(* IEC 61131-3 sources: daoli-st-library/DL_Process (part 46) *)

(* ---- FB_DL_PowderDosingLoss.st ---- *)
// =====================================================================
// FB_DL_PowderDosingLoss.st
// 粉料失重秤增量式配料（皮重→粗给/慢给→落差补偿→稳定结算→学习）
// Loss-in-weight powder dosing FB
// 码位: 16#0005_0458 ~ 16#0005_045C (本件独占 5 槽)
// 修改记录: R29 初版 (按 DISPATCH_R29 序 18)
// =====================================================================
FUNCTION_BLOCK FB_DL_PowderDosingLoss
VAR_INPUT
    bEnable      : BOOL  := FALSE;    // 使能 / Enable
    bStart       : BOOL  := FALSE;    // 上升沿开始一批 / Start batch on edge
    bReset       : BOOL  := FALSE;    // 复位 / Reset
    fWeight_g    : REAL  := 0.0;      // 秤读数 0~500000 g / Scale weight [g]
    fTarget_g    : REAL  := 1000.0;   // 目标投料量 >0 g / Target dose [g]
    fTare_g      : REAL  := 0.0;      // 皮重 ≥0 g / Tare [g]
    fSlowBand_g  : REAL  := 100.0;    // 转慢速余量 >0 g / Slow-down band [g]
    fLead_g      : REAL  := 0.0;      // 落差学习初值 0~500 g / Lead compensation [g]
    fLeadMax_g   : REAL  := 300.0;    // 落差限幅 1~2000 g / Lead limit [g]
    fDevMax_g    : REAL  := 5.0;      // 允许偏差 >0 g / Allowed deviation [g]
    bSlowCmd     : BOOL  := FALSE;    // 慢速输出确认 / Slow feed ack
    tSettleTime  : TIME  := T#500MS;  // 停料稳定时 T#10MS~T#10S / Settle time [s]
    tBatchMax    : TIME  := T#2M;     // 单批超时 T#1S~T#30M / Batch timeout [s]
END_VAR
VAR_OUTPUT
    fNet_g       : REAL;              // 本批净投料 g / Net dosed [g]
    fErr_g       : REAL;              // 本批偏差 g / Deviation [g]
    bDone        : BOOL;              // 批完成（单拍）/ Batch done pulse
    bBusy        : BOOL;              // 配料中 / Busy
    fLeadLearn_g : REAL;              // 更新后落差学习值 g / Learned lead [g]
    eErr         : UDINT;             // 错误码 / Error code
END_VAR
VAR
    rtrigStart   : R_TRIG;            // 启动沿检测（无条件刷新）/ Start edge detector
    tonSettle    : TON;               // 停料稳定定时器（无条件刷新）/ Settle timer
    tonBatch     : TON;               // 单批超时定时器（无条件刷新）/ Batch timeout timer
    fTareSnap_g  : REAL;              // 批开始皮重快照 / Tare snapshot at batch start [g]
    fWeightPrev  : REAL;              // 上拍秤读数快照 / Previous weight snapshot [g]
    fNetNow_g    : REAL;              // 本拍净重 / Net weight this cycle [g]
    fNetStart_g  : REAL;              // 批开始净重基准 / Net baseline at batch start [g]
    fStopPt_g    : REAL;              // 提前停止点（目标-慢带-落差）/ Early stop point [g]
    bFastPhase   : BOOL;              // 高速给料相 / Fast feed phase
    bSettling    : BOOL;              // 停料稳定相 / Settling phase
    tSettleS     : REAL;              // 稳定时秒值 / Settle seconds [s]
    tBatchMaxS   : REAL;              // 批超时秒值 / Batch timeout seconds [s]
    bAbortLatch  : BOOL := FALSE;     // 中止锁存（方向反/超时）/ Abort latch
    xFirstScan   : BOOL  := TRUE;     // 首扫标记 / First-scan flag
END_VAR

// ---------------------------------------------------------------------
// 代码位表（本件独占，勿复用）:
//   16#0005_0458 信息 批完成、偏差在容差内
//   16#0005_0459 故障 秤值非有限 / 皮重为负或超量程 / tSettleTime 非法
//   16#0005_045A 故障 fTarget_g ≤ 0 / fSlowBand_g ≥ fTarget_g / fLeadMax_g ≤ 0（组态错）
//   16#0005_045B 信息 批完成但偏差 > fDevMax_g → 结算照出、落差不学习
//   16#0005_045C 故障 进料期重量上升（方向反）或超 tBatchMax → 中止锁存（方向反优先）
// ---------------------------------------------------------------------

// ---- 时间转秒 / Times to seconds ----
tSettleS := TIME_TO_REAL(tSettleTime) / 1000.0;     // 稳定时秒 / Settle [s]
tBatchMaxS := TIME_TO_REAL(tBatchMax) / 1000.0;     // 批超时秒 / Batch max [s]

// ---- 启动沿检测（无条件刷新）/ Start edge, unconditional ----
rtrigStart(CLK := bStart);      // 沿检测 / Edge detection

// ---- 非有限与皮重闸（故障级）/ Finite and tare gate ----
IF (fWeight_g <> fWeight_g) OR (ABS(fWeight_g) >= 1.0E12)
   OR (fTare_g < 0.0) OR (fTare_g > 500000.0)
   OR (tSettleTime = T#0MS) OR (tSettleS < 0.01) OR (tSettleS > 10.0) THEN
    bBusy := FALSE;             // 停止 / Not busy
    bAbortLatch := TRUE;        // 中止锁存 / Abort latch
    eErr := 16#0005_0459;       // 故障码 / Fault code
    RETURN;                     // 本拍结束 / End of cycle
END_IF

// ---- 组态错闸 / Configuration fault gate ----
IF (fTarget_g <= 0.0) OR (fSlowBand_g >= fTarget_g) OR (fLeadMax_g <= 0.0)
   OR (fDevMax_g <= 0.0)
   OR (tBatchMax = T#0MS) OR (tBatchMaxS < 1.0) OR (tBatchMaxS > 1800.0) THEN
    eErr := 16#0005_045A;       // 故障码 / Fault code
    RETURN;                     // 本拍结束 / End of cycle
END_IF

// ---- 首扫初始化（R16 首扫纪律）/ First-scan initialization ----
IF xFirstScan THEN
    fLeadLearn_g := fLead_g;    // 学习值取初值 / Learn value from init
    fWeightPrev := fWeight_g;   // 快照对齐 / Snapshot align
    bDone := FALSE;             // 脉冲复位 / Pulse reset
    xFirstScan := FALSE;        // 清标记 / Clear flag
END_IF

// ---- 完成脉冲单拍化 / Done pulse one-cycle ----
IF bDone THEN
    bDone := FALSE;             // 下一拍清 / Clear next cycle
END_IF

// ---- 使能撤销 / Disable ----
IF NOT bEnable THEN
    bBusy := FALSE;             // 停止 / Not busy
    bFastPhase := FALSE;        // 粗给退出 / Fast off
    bSettling := FALSE;         // 稳定退出 / Settle off
    eErr := 16#0005_0458;       // 信息级：空闲 / Info: idle
    RETURN;                     // 本拍结束 / End of cycle
END_IF

// ---- 复位：清中止锁存与学习值回初值 / Reset: clear latch, learn back to init ----
IF bReset THEN
    bAbortLatch := FALSE;       // 解锁存 / Release latch
    bBusy := FALSE;             // 停止 / Not busy
    bFastPhase := FALSE;        // 粗给退出 / Fast off
    bSettling := FALSE;         // 稳定退出 / Settle off
    fLeadLearn_g := fLead_g;    // 学习值回初值 / Learn to init
END_IF

// ---- 中止锁存路径 / Abort latch path ----
IF bAbortLatch THEN
    bBusy := FALSE;             // 停止（保留已投量）/ Stopped, dose kept
    eErr := 16#0005_045C;       // 故障码回放 / Fault code replay
    RETURN;                     // 本拍结束 / End of cycle
END_IF

// ---- 每拍净重与方向监控 / Per-cycle net and direction monitor ----
fNetNow_g := fWeight_g - fTare_g;   // 净重 / Net [g]
IF fNetNow_g < 0.0 THEN
    fNetNow_g := 0.0;           // 负值钳 0 / Clamp to 0
    eErr := 16#0005_0459;       // 槽 2 登记 / Slot 2
END_IF

// ---- 启动沿受理（bBusy=FALSE 才受理）/ Accept start edge when idle ----
IF rtrigStart.Q AND (NOT bBusy) THEN
    fTareSnap_g := fTare_g;     // 皮重快照 / Tare snapshot
    fNetStart_g := fNetNow_g;   // 净重基准 / Net baseline
    fWeightPrev := fWeight_g;   // 快照对齐 / Snapshot align
    fStopPt_g := fTarget_g - fSlowBand_g - fLeadLearn_g;    // 提前停止点含落差 / Stop point with lead
    IF fStopPt_g < 0.0 THEN
        fStopPt_g := 0.0;       // 防负停止点 / Guard negative stop
    END_IF
    bBusy := TRUE;              // 配料中 / Busy
    bFastPhase := TRUE;         // 粗给开始 / Fast feed
    bSettling := FALSE;         // 非稳定相 / Not settling
END_IF

// ---- 批运行路径 / Batch active path ----
IF bBusy THEN
    // 单批超时监控 / Batch timeout monitor
    tonBatch(IN := bBusy, PT := tBatchMax);     // 无条件刷新 / Unconditional refresh

    // 方向监控：进料期重量上升 → 方向反（根因优先，先于超时判）/ Direction: rising weight fault first
    IF fWeight_g > (fWeightPrev + 1.0) THEN
        bAbortLatch := TRUE;    // 中止锁存 / Abort latch
        bBusy := FALSE;         // 停止 / Not busy
        bFastPhase := FALSE;    // 粗给退出 / Fast off
        bSettling := FALSE;     // 稳定退出 / Settle off
        eErr := 16#0005_045C;   // 故障码：方向反 / Fault code: reversed
        fWeightPrev := fWeight_g;   // 快照对齐 / Align snapshot
        RETURN;                 // 本拍结束 / End of cycle
    END_IF

    // 批超时（方向反已优先返回）/ Batch timeout after direction check
    IF tonBatch.Q THEN
        bAbortLatch := TRUE;    // 中止锁存 / Abort latch
        bBusy := FALSE;         // 停止（保留已投量）/ Stopped, dose kept
        bFastPhase := FALSE;    // 粗给退出 / Fast off
        bSettling := FALSE;     // 稳定退出 / Settle off
        eErr := 16#0005_045C;   // 故障码：超时 / Fault code: timeout
        RETURN;                 // 本拍结束 / End of cycle
    END_IF

    // ---- 给料相控制 / Feed phase control ----
    IF bFastPhase THEN
        // 高速粗给：净投量未达提前停止点 / Fast: below stop point
        IF (fNetNow_g - fNetStart_g) >= fStopPt_g THEN
            bFastPhase := FALSE;    // 转慢速精给 / To slow feed
        END_IF
        // 慢速转换确认（bSlowCmd 为外部确认，此处登记不强制）/ Slow ack registered externally
    END_IF

    // 停料判定：慢给相已达目标（含落差提前）/ Stop: reached target with lead
    IF (NOT bFastPhase) AND ((fNetNow_g - fNetStart_g) >= (fTarget_g - fLeadLearn_g)) THEN
        bSettling := TRUE;      // 停料稳定相 / Settling
        tonSettle(IN := TRUE, PT := tSettleTime);   // 稳定计时 / Settle timing
    END_IF

    // ---- 稳定后结算 / Settle then finalize ----
    IF bSettling THEN
        tonSettle(IN := TRUE, PT := tSettleTime);   // 无条件刷新 / Unconditional refresh
        IF tonSettle.Q THEN
            fNet_g := fNetNow_g - fNetStart_g;  // 结算净投量 / Finalize net
            fErr_g := fNet_g - fTarget_g;       // 偏差 / Deviation
            bDone := TRUE;      // 完成脉冲 / Done pulse
            bBusy := FALSE;     // 停止 / Not busy
            bSettling := FALSE; // 稳定退出 / Settle off
            IF ABS(fErr_g) <= fDevMax_g THEN
                // 落差学习：LIMIT(0, fLead + 0.5×fErr, fLeadMax)，0.5 阻尼防振荡
                // Lead learning: LIMIT with 0.5 damping factor
                fLeadLearn_g := fLeadLearn_g + 0.5 * fErr_g;    // 学习更新 / Learn update
                IF fLeadLearn_g < 0.0 THEN
                    fLeadLearn_g := 0.0;    // 下限 / Lower limit
                ELSIF fLeadLearn_g > fLeadMax_g THEN
                    fLeadLearn_g := fLeadMax_g;     // 上限 / Upper limit
                END_IF
                eErr := 16#0005_0458;   // 信息级：批完成 / Info: done
            ELSE
                eErr := 16#0005_045B;   // 信息级：超差结算不学习 / Info: no learning
            END_IF
        END_IF
    END_IF
ELSE
    tonBatch(IN := FALSE, PT := tBatchMax);     // 定时器复位 / Timer reset
    tonSettle(IN := FALSE, PT := tSettleTime);  // 定时器复位 / Timer reset
END_IF

// ---- 上拍快照更新 / Previous snapshot update ----
fWeightPrev := fWeight_g;       // 快照 / Snapshot

END_FUNCTION_BLOCK

(* ---- FB_DL_PressFitCurveArchive.st ---- *)
(*
  Component : FB_DL_PressFitCurveArchive
  Category  : DL_Process
  Type      : FB
  Version   : 1.0.0
  CodeSeg   : 16#06_0_3B
  Summary   : 压装曲线特征点归档与批次追溯：四特征点环形缓存按批次号索引，R_TRIG 沿触发归档。
              Press-fit curve feature archive by batch index in a ring buffer, triggered on a rising edge.
  溯源声明  : 道莅自研 clean-room
  边界安全  : 批次号域闸（> 0，防非法索引）；环形缓冲下标 1..NMAX 硬界，写前钳制防越界；
              特征点非有限（NaN 自反 + Inf 上限）拦截；查询命中用整数相等（DINT）；
              R_TRIG 每拍无条件刷新（段 0）；缓冲满环回写并置 bWrapped 提示；计数防回卷。
  复用      : 无
*)

FUNCTION_BLOCK FB_DL_PressFitCurveArchive
VAR_INPUT
    bRun       : BOOL;                  (* 归档使能 · Enable *)
    bArchCmd   : BOOL;                  (* 归档指令 [事件]，沿触发 · Archive command, edge *)
    nBatchNo   : DINT;                  (* 批次号 [号]，域 > 0 · Batch number *)
    fF1KN      : LREAL;                 (* 特征点 1：起步压力 [kN] · Feature 1 onset force *)
    fF2MM      : LREAL;                 (* 特征点 2：起步位移 [mm] · Feature 2 onset travel *)
    fF3KN      : LREAL;                 (* 特征点 3：峰值压力 [kN] · Feature 3 peak force *)
    fF4MM      : LREAL;                 (* 特征点 4：终点位移 [mm] · Feature 4 end travel *)
    nQueryNo   : DINT;                  (* 追溯查询批次号 [号] · Query batch number *)
    fEps       : LREAL := 1.0E-6;       (* 浮点判零容差 [实数域] · Floating zero tolerance *)
END_VAR
VAR_OUTPUT
    bArchOk  : BOOL;                    (* 本拍归档成功 [开关] · Archive succeeded this scan *)
    bWrapped : BOOL;                    (* 环已回卷覆盖标志 · Ring wrapped flag *)
    bFound   : BOOL;                    (* 查询命中标志 · Query hit flag *)
    fQ1KN    : LREAL;                   (* 查询特征 1 [kN] · Queried feature 1 *)
    fQ2MM    : LREAL;                   (* 查询特征 2 [mm] · Queried feature 2 *)
    fQ3KN    : LREAL;                   (* 查询特征 3 [kN] · Queried feature 3 *)
    fQ4MM    : LREAL;                   (* 查询特征 4 [mm] · Queried feature 4 *)
    nUsed    : INT;                     (* 环内已用槽数 [槽] · Used slots *)
    bError   : BOOL;                    (* 故障标志，与故障码配对 · Fault flag paired with codes *)
    uErrorId : UDINT;                   (* 事件码 16#0000_003B，0 无事件 · Event code *)
END_VAR
VAR
    uCode   : WORD;     (* 码位暂存，每拍重算 [码] · Code staging *)
    rTrigArc: R_TRIG;   (* 归档上升沿，每拍无条件刷新 · Archive edge detection *)
    aIdx    : ARRAY[1..8] OF DINT;      (* 批次号索引槽 [号] · Batch index slots *)
    aF1     : ARRAY[1..8] OF LREAL;     (* 特征 1 缓存 [kN] · Feature 1 buffer *)
    aF2     : ARRAY[1..8] OF LREAL;     (* 特征 2 缓存 [mm] · Feature 2 buffer *)
    aF3     : ARRAY[1..8] OF LREAL;     (* 特征 3 缓存 [kN] · Feature 3 buffer *)
    aF4     : ARRAY[1..8] OF LREAL;     (* 特征 4 缓存 [mm] · Feature 4 buffer *)
    nHead   : INT;      (* 环形写头下标 [索引] · Ring head index *)
    nI      : INT;      (* 查询循环下标 [索引] · Query loop index *)
    bSigOk  : BOOL;     (* 输入有效标志 · Input validity flag *)
    nCycles : UDINT;    (* 归档累计 [次]，防回卷 · Archive count *)
END_VAR
VAR CONSTANT
    DL_PCA_NMAX : INT := 8;             (* 环形缓冲容量 [槽] · Ring capacity *)
    DL_PCA_WRAP : UDINT := 4294967290;  (* 计数防回卷余量 [次] · Counter wrap guard *)
END_VAR

(* === 段 0 · 实例刷新（每拍无条件，红线 7）=== *)
IF nHead < 1 THEN
    nHead := 1;                         (* 写头初值钳 1，防数组零下标越界 / Clamp the head to one *)
END_IF
rTrigArc(CLK := bArchCmd);              (* 归档沿检测 / Archive edge *)

(* === 段 1 · 输入校验与量程闸 === *)
uCode := 16#0000;                       // 每拍清码（可达清零基线）/ Clear codes each scan
bSigOk := (nBatchNo > 0)                                             // 批次号正域闸 / Batch number gate
          AND (fF1KN = fF1KN) AND (fF2MM = fF2MM)                     // 特征点非有限拦截 / Non-finite guards
          AND (fF3KN = fF3KN) AND (fF4MM = fF4MM)
          AND (ABS(fF1KN) < 1.0E308) AND (ABS(fF3KN) < 1.0E308)       // Inf 上限判据 / Inf limits
          AND (ABS(fF2MM) < 1.0E308) AND (ABS(fF4MM) < 1.0E308)
          AND (fF3KN > fF1KN);                                        // 峰值起步序闸 / Peak above onset
IF NOT bSigOk THEN
    uCode := 16#003B;                   // 故障级：域外，归档拒绝 / Fault: domain invalid
END_IF

(* === 段 2 · 主逻辑：环形归档与批次追溯 === *)
bArchOk := FALSE;                       (* 归档成功标志单拍重建 / Rebuild the success flag *)
IF rTrigArc.Q AND bRun THEN
    IF bSigOk THEN
        aIdx[nHead] := nBatchNo;        (* 写批次索引（头下标受 NMAX 硬界）/ Write the index *)
        aF1[nHead] := fF1KN;            (* 写特征 1 [kN] / Write feature 1 *)
        aF2[nHead] := fF2MM;            (* 写特征 2 [mm] / Write feature 2 *)
        aF3[nHead] := fF3KN;            (* 写特征 3 [kN] / Write feature 3 *)
        aF4[nHead] := fF4MM;            (* 写特征 4 [mm] / Write feature 4 *)
        bArchOk := TRUE;                (* 归档成功 / Archive done *)
        IF nUsed < DL_PCA_NMAX THEN
            nUsed := nUsed + 1;         (* 未满先增用量 / Grow usage *)
        ELSE
            bWrapped := TRUE;           (* 满环回卷提示 / Ring wrapped flag *)
        END_IF
        nHead := (nHead MOD DL_PCA_NMAX) + 1;   (* 写头循环推进，界内 / Advance the head in bounds *)
        IF nCycles < DL_PCA_WRAP THEN
            nCycles := nCycles + 1;     (* 归档计数 / Count archives *)
        END_IF
    END_IF
END_IF
(* 追溯查询：按批次号线性匹配（DINT 等值合法）/ Trace query by batch number *)
bFound := FALSE;                        (* 命中标志单拍重建 / Rebuild the hit flag *)
IF (nQueryNo > 0) AND (nUsed >= 1) THEN
    FOR nI := 1 TO DL_PCA_NMAX DO
        IF nI <= nUsed THEN
            IF aIdx[nI] = nQueryNo THEN
                fQ1KN := aF1[nI];       (* 命中回放特征 1 [kN] / Replay feature 1 *)
                fQ2MM := aF2[nI];       (* 回放特征 2 [mm] / Replay feature 2 *)
                fQ3KN := aF3[nI];       (* 回放特征 3 [kN] / Replay feature 3 *)
                fQ4MM := aF4[nI];       (* 回放特征 4 [mm] / Replay feature 4 *)
                bFound := TRUE;         (* 命中 / Hit *)
                EXIT;                   (* 单命中即止 / Stop on first hit *)
            END_IF
        END_IF
    END_FOR
END_IF

(* === 段 3 · 输出映射与故障码 === *)
IF NOT bFound THEN
    fQ1KN := 0.0;                       (* 未命中输出安全零（哨兵）/ Safe zeros on miss *)
    fQ2MM := 0.0;
    fQ3KN := 0.0;
    fQ4MM := 0.0;
END_IF
IF NOT bRun THEN
    bWrapped := FALSE;                  (* 撤使能清回卷提示（可达清零）/ Clear on disable *)
END_IF
bError := (uCode <> 16#0000);           (* 故障标志配对 / Fault flag paired *)
uErrorId := WORD_TO_UDINT(uCode);       (* 码位单点写入（16#0000_003B 形态）/ Single write point *)
END_FUNCTION_BLOCK

(* ---- FB_DL_PrintRegisterAutoTrimSeq.st ---- *)
(*
  DL Factory R83 | FB_DL_PrintRegisterAutoTrimSeq
  功能：印刷套准自动调整状态机，横纵套准误差超差后按三级阶梯逐级小步修正，每步等稳定窗后复评，超步数上限锁故障码。
  开源溯源：无（clean-room 自研，依据公开工艺公式，来源=行业通用公式，许可证=MIT，借鉴点=公式结构）
  规则：R1-R21 全遵守
  ------------------------------------------------------------------
  分类 DL_Process ｜ 复杂度 cx4 ｜ 版本 v1.0.0 ｜ 平台 纯 IEC 61131-3（TON、R_TRIG、LREAL）
  边界：一 只出三级修正命令，不驱动版辊电机本体、不做套准标记识别（识别归前级视觉件属主）；
        二 阶梯次序固定：一 色标偏移（管横向）→ 二 版辊相位（管纵向）→ 三 张力微调（管纵向残差）；
           一与二同属偏移域共用 eVern 相、由 _nLadder 区分下发通道；三独立占 eTens 相（力值量禁与长度量混加）；
        三 每步下发后等回执沿（脉冲语义，须回零后再置位），否则超时锁 104；每相只允许一个专属定时器，
           IN 只串本相使能与锁存闸，相迁移即 IN 归假并自复位（R18）；tonVern 与 tonTens 分属互斥相、
           无同拍双窗，故 R100 配比约束不适用；
        四 小步下发前方向分列（偏正 ｜ 偏负各占一分支，R146），下发后立即饱和到本通道限值；
        五 命令累加量在复位沿保持末值（已下发修正不得被复位抹掉），作用域在段 1 逐项声明；
           无全局变量、无外部变量声明、无物理地址寻址。
  量纲自检：长度量 [mm] 通道 = fErrCross / fTolCross / fStepVernier / fCmdLimit 与 fErrMachine / fTolMachine / fStepPhase；
        力值量 [N] 通道 = fStepTension / fTensLimit（禁与长度量相加）；组态闸另校各步长落在本通道限值内防越窗振荡。
  输出契约：三级命令为累加型且已饱和；bDone 为电平保持位（新循环起点同拍清零，R28 5.9）；iErrCode 为锁存回放，故障锁存唯一解除路径为 bReset 上升沿（R188）。
  修订记录：2026-11-24 v1.0.0 R83 首版（批 R83 · 序号 37）
*)

TYPE E_DL_PraPhase :
(
    eIdle   := 0,  // 空闲等启动沿 / idle, waiting for the start edge
    eEval   := 10, // 评估：判容差选阶梯并下发（单拍相）/ evaluate, judge and issue in one scan
    eVern   := 20, // 偏移修正等回执（承载阶梯一二）/ offset trim, waiting for the acknowledgement
    eTens   := 30, // 张力修正等回执（承载阶梯三）/ tension trim, waiting for the acknowledgement
    eSettle := 40, // 稳定等稳定窗 / settling, waiting for the window
    eDone   := 50, // 完成：误差在容差内 / done, the error is inside the tolerance
    eFault  := 90  // 故障：成因锁存等复位沿 / fault, the cause is latched until the reset edge
);
END_TYPE

TYPE E_DL_PraCause :
(
    eNone      := 0, // 无成因 / no cause
    eCfgBad    := 1, // 组态越域或量纲失配（故障级，与 bError 配对）/ configuration out of domain, fault grade paired with bError
    eNotFinite := 2, // 入参非有限 NaN 或 Inf（故障级，与 bError 配对）/ non-finite input, fault grade paired with bError
    eStepLimit := 3, // 步数上限耗尽仍超差（故障级，与 bError 配对）/ step budget exhausted, fault grade paired with bError
    eAckTo     := 4, // 步进回执超时（故障级，与 bError 配对）/ acknowledgement timeout, fault grade paired with bError
    ePhaseBad  := 5  // 非法相位兜底（故障级，与 bError 配对）/ illegal phase fallback, fault grade paired with bError
);
END_TYPE

FUNCTION_BLOCK FB_DL_PrintRegisterAutoTrimSeq
VAR CONSTANT
    DL_PRA_LADDER_VERN   : INT := 1; // 阶梯一：色标偏移通道 [级] / ladder one, the register mark offset channel [stage]
    DL_PRA_LADDER_PHASE  : INT := 2; // 阶梯二：版辊相位通道 [级] / ladder two, the plate cylinder phase channel [stage]
    DL_PRA_LADDER_TENS   : INT := 3; // 阶梯三：张力微调通道 [级] / ladder three, the tension trim channel [stage]
    DL_PRA_PHASE_TRY_MAX : INT := 2; // 阶梯二连续复用预算，超限升阶梯三 [次] / the reuse budget of ladder two [time]
END_VAR
VAR_INPUT
    bEnable      : BOOL := TRUE;   // 使能，失能退回空闲（命令保持末值）[-] / enable, a disable returns to idle holding the commands
    bReset       : BOOL := FALSE;  // 复位上升沿清故障锁存与步数 [-]/ reset rising edge clears the latch and the steps
    bStart       : BOOL := FALSE;  // 启动电平，上升沿起一轮调整 [-]/ start level, its rising edge begins one round
    bStepAck     : BOOL := FALSE;  // 步进执行回执（脉冲语义须回零）[-]/ the step acknowledgement, pulse semantics
    fErrCross    : LREAL := 0.0;   // 横向套准误差（正 = 偏大）[mm] / the cross register error, positive means too large [mm]
    fErrMachine  : LREAL := 0.0;   // 纵向套准误差（正 = 偏大）[mm] / the machine register error, positive means too large [mm]
    fTolCross    : LREAL := 0.10;  // 横向容差半带宽 [mm] / the cross tolerance half band [mm]
    fTolMachine  : LREAL := 0.10;  // 纵向容差半带宽 [mm] / the machine tolerance half band [mm]
    fStepVernier : LREAL := 0.05;  // 色标偏移单步量（阶梯一）[mm] / the offset step of ladder one [mm]
    fStepPhase   : LREAL := 0.05;  // 版辊相位单步等效位移（阶梯二）[mm] / the phase step of ladder two [mm]
    fStepTension : LREAL := 2.0;   // 张力微调单步量（阶梯三）[N] / the tension step of ladder three [N]
    fCmdLimit    : LREAL := 5.0;   // 长度通道命令饱和限（对称）[mm] / the symmetric length channel command limit [mm]
    fTensLimit   : LREAL := 200.0; // 张力通道命令饱和限（对称）[N] / the symmetric tension channel command limit [N]
    nMaxStep     : INT := 20;      // 单轮步数上限 [步] / the step budget of one round [step]
    tSettle      : TIME := T#2S;   // 单步后稳定窗 [毫秒] / the settling window after each step [millisecond]
    tAckTo       : TIME := T#10S;  // 步进回执超时窗 [毫秒] / the acknowledgement timeout [millisecond]
END_VAR
VAR_OUTPUT
    bBusy       : BOOL := FALSE;   // 本轮调整进行中 [-] / the round is in progress
    bDone       : BOOL := FALSE;   // 到达容差（保持式，新循环起点清零）[-] / reached the tolerance, held until a new round
    bFault      : BOOL := FALSE;   // 故障锁存 [-] / the fault latch
    bError      : BOOL := FALSE;   // 故障标志，与锁存位同源 [-] / the fault flag sharing the latch source
    iErrCode    : INT := 0;        // 错误码（锁存回放，复位沿清零）[码] / the error code replayed from the latch [code]
    ePhase      : E_DL_PraPhase := E_DL_PraPhase.eIdle; // 相位出口 [枚举] / the phase outlet [enum]
    fVernierOut : LREAL := 0.0;    // 色标偏移命令（累加已饱和）[mm] / the offset command, accumulated [mm]
    fPhaseOut   : LREAL := 0.0;    // 版辊相位命令（累加已饱和）[mm] / the phase command, accumulated [mm]
    fTensionOut : LREAL := 0.0;    // 张力微调命令（累加已饱和）[N] / the tension command, accumulated [N]
    nStepUsed   : INT := 0;        // 本轮已执行步数 [步] / the executed step count [step]
    nLadderIdx  : INT := 1;        // 当前阶梯编号（诊断 1/2/3）[级] / the current ladder index for diagnostics [stage]
    bInTol      : BOOL := FALSE;   // 横纵误差均在容差内 [-] / both errors are inside the tolerance
    bStepActive : BOOL := FALSE;   // 某级小步正在等回执 [-] / a step is waiting for the acknowledgement
END_VAR
VAR
    rtStart   : R_TRIG; // 启动沿，段 0 无条件刷新 / the start edge, refreshed unconditionally
    rtReset   : R_TRIG; // 复位沿，段 0 无条件刷新 / the reset edge, refreshed unconditionally
    rtAck     : R_TRIG; // 回执沿，段 0 无条件刷新 / the acknowledgement edge, refreshed unconditionally
    tonVern   : TON;    // 偏移回执超时窗，段 0 无条件刷新 / the offset acknowledgement timeout
    tonTens   : TON;    // 张力回执超时窗，段 0 无条件刷新 / the tension acknowledgement timeout
    tonSettle : TON;    // 稳定窗，段 0 无条件刷新 / the settling window
    _ePhase   : E_DL_PraPhase := E_DL_PraPhase.eIdle; // 内部相位，CASE 唯一写入目标 / the internal phase, the only CASE target
    _eCause   : E_DL_PraCause := E_DL_PraCause.eNone; // 故障级成因，锁存至复位沿 / the fault cause latched until reset
    _bFault   : BOOL := FALSE; // 故障锁存位 [-] / the fault latch
    _bReq     : BOOL := FALSE; // 本拍故障请求（单拍预清，R107）[-] / the scan fault request, pre-cleared
    _iErrTmp  : INT := 0;      // 本拍码位暂存 [码] / the scan code [code]
    _iErrLch  : INT := 0;      // 码位锁存槽 [码] / the latched code [code]
    _bDone    : BOOL := FALSE; // 完成位内部锁存（清零归属：段 1 复位沿与段 2 启动沿）[-] / the internal done bit
    _bInit    : BOOL := FALSE; // 首扫初始化完成标志（R310）[-] / the first scan initialisation flag
    _bCfgOk   : BOOL := FALSE; // 组态参数域内 [-] / the configuration is inside the domain
    _bFinOk   : BOOL := FALSE; // 全部浮点入参有限 [-] / every floating input is finite
    _bInTol   : BOOL := FALSE; // 容差判据原始值 [-] / the raw tolerance verdict
    _nLadder  : INT := 1;      // 当前阶梯编号 1/2/3 [级] / the current ladder index [stage]
    _nTry     : INT := 0;      // 阶梯二连续使用次数 [次] / the consecutive uses of ladder two [time]
    _nStep    : INT := 0;      // 已执行步数累计 [步] / the executed step count [step]
    _fVernAcc : LREAL := 0.0;  // 偏移命令累加量（复位保持末值）[mm] / the offset accumulator held across a reset [mm]
    _fPhaseA  : LREAL := 0.0;  // 相位命令累加量（复位保持末值）[mm] / the phase accumulator held across a reset [mm]
    _fTensAcc : LREAL := 0.0;  // 张力命令累加量（复位保持末值）[N] / the tension accumulator held across a reset [N]
END_VAR
// 段 0｜定时器与沿检测无条件周期刷新，IN 只串本相使能与锁存闸，禁 R_TRIG.Q 直连（R7 / R18 / FB50-1）
rtStart(CLK := bStart); // 启动沿无条件刷新 / unconditional refresh of the start edge
rtReset(CLK := bReset); // 复位沿无条件刷新 / unconditional refresh of the reset edge
rtAck(CLK := bStepAck); // 回执沿无条件刷新 / unconditional refresh of the acknowledgement edge
tonVern(IN := (_ePhase = E_DL_PraPhase.eVern) AND (NOT _bFault), PT := tAckTo); // 偏移回执超时窗，只串 eVern 相 / the offset timeout gated by eVern only
tonTens(IN := (_ePhase = E_DL_PraPhase.eTens) AND (NOT _bFault), PT := tAckTo); // 张力回执超时窗，只串 eTens 相 / the tension timeout gated by eTens only
tonSettle(IN := (_ePhase = E_DL_PraPhase.eSettle) AND (NOT _bFault), PT := tSettle); // 稳定窗，只串 eSettle 相 / the settling window gated by eSettle only

// 段 1｜首扫初始化与复位沿同块，作用域逐项声明（R310 / R311，两者初始化项同款）
IF (NOT _bInit) OR rtReset.Q THEN // 首扫一拍或复位沿 / the first scan or the reset edge
    _bInit := TRUE; // 首扫完成标志（复位沿重复置位同效）/ the first scan flag, the same effect on reset
    _bFault := FALSE; // 作用域一：清故障锁存位 / scope one, clear the fault latch
    _eCause := E_DL_PraCause.eNone; // 作用域一：清故障级成因 / scope one, clear the fault cause
    _iErrLch := 0; // 作用域一：清码位锁存槽 / scope one, clear the code slot
    _bDone := FALSE; // 作用域二：清完成位（电平保持位由复位沿解除）/ scope two, clear the held done bit
    _ePhase := E_DL_PraPhase.eIdle; // 作用域二：迁回空闲相 / scope two, migrate back to idle
    _nStep := 0; // 作用域三：清累计步数 / scope three, clear the accumulated steps
    _nLadder := DL_PRA_LADDER_VERN; // 作用域三：阶梯回到一 / scope three, the ladder returns to one
    _nTry := 0; // 作用域三：清阶梯二使用次数 / scope three, clear the ladder two counter
END_IF // 作用域之外的保持项：_fVernAcc ｜ _fPhaseA ｜ _fTensAcc 三项保持末值（已下发修正不得被复位抹掉）
// 段 2｜启动沿：新循环起点同拍清完成位与步数（R28 5.9 清零点）
IF rtStart.Q THEN // 启动沿 / the start edge
    _bDone := FALSE; // 完成位清零（上一轮遗留）/ clear the done bit left by the previous round
    _nStep := 0; // 步数清零 / clear the step count
    _nLadder := DL_PRA_LADDER_VERN; // 阶梯回到一 / the ladder returns to one
    _nTry := 0; // 阶梯二使用次数清零 / clear the ladder two counter
END_IF
// 段 3｜组态域闸：参与判据换算的引脚逐项枚举，含量纲尺度自检（R151 / R20 / R272）
_bCfgOk := (fTolCross > 0.0) AND (fTolMachine > 0.0) AND (fCmdLimit > 0.0) AND (fTensLimit > 0.0) // 容差与两通道饱和限须为正 / the tolerances and both channel limits must be positive
    AND (fStepVernier > 0.0) AND (fStepVernier <= fCmdLimit) // 阶梯一步长正且在限内 / ladder one step positive and inside its limit
    AND (fStepPhase > 0.0) AND (fStepPhase <= fCmdLimit) // 阶梯二步长正且在限内 / ladder two step positive and inside its limit
    AND (fStepTension > 0.0) AND (fStepTension <= fTensLimit) // 阶梯三步长正且在限内 / ladder three step positive and inside its limit
    AND (nMaxStep >= 1) AND (tSettle > T#0S) AND (tAckTo > T#0S); // 步数预算与两个时间引脚域闸 / the step budget and the time gates
// 段 4｜非有限闸：9 个浮点入参显式全枚举，NaN 与 Inf 双拦截（R21 / R272）
_bFinOk := (fErrCross > -1.0E30) AND (fErrCross < 1.0E30) AND (fErrMachine > -1.0E30) AND (fErrMachine < 1.0E30) // 横纵误差有限 / both register errors are finite
    AND (fTolCross > -1.0E30) AND (fTolCross < 1.0E30) AND (fTolMachine > -1.0E30) AND (fTolMachine < 1.0E30) // 横纵容差有限 / both tolerances are finite
    AND (fStepVernier > -1.0E30) AND (fStepVernier < 1.0E30) AND (fStepPhase > -1.0E30) AND (fStepPhase < 1.0E30) // 阶梯一二步长有限 / the ladder one and two steps are finite
    AND (fStepTension > -1.0E30) AND (fStepTension < 1.0E30) // 阶梯三步长有限 / the ladder three step is finite
    AND (fCmdLimit > -1.0E30) AND (fCmdLimit < 1.0E30) AND (fTensLimit > -1.0E30) AND (fTensLimit < 1.0E30); // 两通道限值有限 / both channel limits are finite
// 段 5｜容差实时判据：两侧均须满足，且组态与有限性闸位同时成立
_bInTol := _bFinOk AND _bCfgOk AND (ABS(fErrCross) <= fTolCross) AND (ABS(fErrMachine) <= fTolMachine); // 双闸位与双容差同真 / both gates and both tolerances hold
// 段 6｜故障判据与锁存：请求位每拍预清，锁存与迁相同拍执行（R107 / FB50-1④ / R152）
_bReq := FALSE; // 单拍请求位预清（不含 Prev 快照与锁存量）/ pre-clear the single scan request
_iErrTmp := 0; // 本拍码位暂存预清 / pre-clear the scan code
IF (NOT _bFault) AND (NOT _bCfgOk) THEN // 组态越域 / the configuration is out of domain
    _eCause := E_DL_PraCause.eCfgBad; _iErrTmp := 101; // 故障级成因与码位：组态越域 / fault cause and code, the configuration is out of domain
    bError := TRUE; // R45 配对：故障级码位同拍置故障标志 / the fault flag paired with the code
    _bReq := TRUE; // 请求本拍锁存 / request the latch
END_IF
IF (NOT _bFault) AND (NOT _bFinOk) THEN // 入参非有限 / a non-finite input
    _eCause := E_DL_PraCause.eNotFinite; _iErrTmp := 102; // 故障级成因与码位：入参非有限 / fault cause and code, a non-finite input
    bError := TRUE; // R45 配对：故障级码位同拍置故障标志 / the fault flag paired with the code
    _bReq := TRUE; // 请求本拍锁存 / request the latch
END_IF
IF _bReq AND (NOT _bFault) THEN // 锁存只认当拍首因 / latch only the first cause of this scan
    _iErrLch := _iErrTmp; // 码位进锁存槽 / the code enters the latch slot
    _bFault := TRUE; // 置故障锁存位 / raise the fault latch
    _ePhase := E_DL_PraPhase.eFault; // 锁存同拍迁故障相 / migrate to the fault phase in the same scan
END_IF
// 段 7｜相位状态机：ENUM + CASE + ELSE 非法相位兜底（R6 / R128），相内锁存与迁相同分支（FB50-1④）
CASE _ePhase OF
E_DL_PraPhase.eIdle: // 空闲相：退出条件二（启动沿生效 ｜ 使能未给则驻留等下一沿）
    IF bEnable AND rtStart.Q THEN // 启动沿且使能 / the start edge while enabled
        _ePhase := E_DL_PraPhase.eEval; // 迁评估相（拍 N 进入：本相起点 ｜ 本拍行为：拒绝下发 ｜ 拍 N+1 转出：决策相）
    END_IF
E_DL_PraPhase.eEval: // 评估相：单拍决策——判容差、判步数、选阶梯、下发小步
    IF _bInTol THEN // 误差已入容差 / the errors are inside
        _bDone := TRUE; _ePhase := E_DL_PraPhase.eDone; // 置完成位（保持至新循环起点）并迁完成相 / raise done and migrate
    ELSIF _nStep >= nMaxStep THEN // 步数预算耗尽仍超差 / the budget is exhausted
        _eCause := E_DL_PraCause.eStepLimit; _iErrLch := 103; // 故障级成因与码位：步数耗尽 / fault cause and code, the step budget exhausted
        bError := TRUE; // R45 配对：故障级成因同拍置故障标志 / the fault flag paired with the cause
        _bFault := TRUE; _ePhase := E_DL_PraPhase.eFault; // 置锁存并迁故障相 / latch and migrate to the fault phase
    ELSIF (ABS(fErrCross) > fTolCross) THEN // 横向超差：走阶梯一（色标偏移）/ the cross error is out, take ladder one
        _nLadder := DL_PRA_LADDER_VERN; _nTry := 0; // 阶梯登记为一并清阶梯二计数 / register ladder one and clear the counter
        IF fErrCross > 0.0 THEN _fVernAcc := _fVernAcc - fStepVernier; ELSE _fVernAcc := _fVernAcc + fStepVernier; END_IF // 方向分列：偏正减步长 ｜ 偏负加步长 / direction split by the error sign
        IF _fVernAcc > fCmdLimit THEN _fVernAcc := fCmdLimit; ELSIF _fVernAcc < (0.0 - fCmdLimit) THEN _fVernAcc := (0.0 - fCmdLimit); END_IF // 双向饱和到通道限 / two sided saturation
        _nStep := _nStep + 1; _ePhase := E_DL_PraPhase.eVern; // 计一步并迁偏移修正相等回执 / count the step and wait for the acknowledgement
    ELSIF (ABS(fErrMachine) > fTolMachine) AND (_nTry < DL_PRA_PHASE_TRY_MAX) THEN // 纵向超差且阶梯二在预算内 / the machine error is out within the ladder two budget
        _nLadder := DL_PRA_LADDER_PHASE; _nTry := _nTry + 1; // 阶梯登记为二并计一次使用 / register ladder two and count one use
        IF fErrMachine > 0.0 THEN _fPhaseA := _fPhaseA - fStepPhase; ELSE _fPhaseA := _fPhaseA + fStepPhase; END_IF // 相位方向分列 / the phase direction split
        IF _fPhaseA > fCmdLimit THEN _fPhaseA := fCmdLimit; ELSIF _fPhaseA < (0.0 - fCmdLimit) THEN _fPhaseA := (0.0 - fCmdLimit); END_IF // 双向饱和到通道限 / two sided saturation
        _nStep := _nStep + 1; _ePhase := E_DL_PraPhase.eVern; // 计一步并迁偏移修正相等回执 / count the step and wait for the acknowledgement
    ELSE // 纵向超差且阶梯二预算耗尽：升阶梯三（张力微调）/ the budget is gone, escalate to ladder three
        _nLadder := DL_PRA_LADDER_TENS; // 阶梯登记为三 / register ladder three
        IF fErrMachine > 0.0 THEN _fTensAcc := _fTensAcc + fStepTension; ELSE _fTensAcc := _fTensAcc - fStepTension; END_IF // 偏正升张力 ｜ 偏负降张力 / raise the tension when the error is positive
        IF _fTensAcc > fTensLimit THEN _fTensAcc := fTensLimit; ELSIF _fTensAcc < (0.0 - fTensLimit) THEN _fTensAcc := (0.0 - fTensLimit); END_IF // 双向饱和到通道限 / two sided saturation
        _nStep := _nStep + 1; _ePhase := E_DL_PraPhase.eTens; // 计一步并迁张力修正相等回执 / count the step and wait for the acknowledgement
    END_IF
E_DL_PraPhase.eVern: // 偏移修正相：退出条件三（回执沿 ｜ 回执超时 ｜ 使能丢失），本拍事件优先于超时（R275）
    IF NOT bEnable THEN // 使能丢失 / the enable was lost
        _ePhase := E_DL_PraPhase.eIdle; // 退回空闲（命令保持末值）/ back to idle holding the commands
    ELSIF rtAck.Q THEN // 回执沿先消化 / digest the acknowledgement first
        _ePhase := E_DL_PraPhase.eSettle; // 迁稳定相 / migrate to settle
    ELSIF tonVern.Q THEN // 回执超时 / the acknowledgement timed out
        _eCause := E_DL_PraCause.eAckTo; _iErrLch := 104; // 故障级成因与码位：回执超时 / fault cause and code, the acknowledgement timeout
        bError := TRUE; // R45 配对：故障级成因同拍置故障标志 / the fault flag paired with the cause
        _bFault := TRUE; _ePhase := E_DL_PraPhase.eFault; // 置锁存并迁故障相 / latch and migrate to the fault phase
    END_IF
E_DL_PraPhase.eTens: // 张力修正相：退出条件三（回执沿 ｜ 回执超时 ｜ 使能丢失），本拍事件优先于超时（R275）
    IF NOT bEnable THEN // 使能丢失 / the enable was lost
        _ePhase := E_DL_PraPhase.eIdle; // 退回空闲（命令保持末值）/ back to idle holding the commands
    ELSIF rtAck.Q THEN // 回执沿先消化 / digest the acknowledgement first
        _ePhase := E_DL_PraPhase.eSettle; // 迁稳定相 / migrate to settle
    ELSIF tonTens.Q THEN // 回执超时 / the acknowledgement timed out
        _eCause := E_DL_PraCause.eAckTo; _iErrLch := 104; // 故障级成因与码位：回执超时 / fault cause and code, the acknowledgement timeout
        bError := TRUE; // R45 配对：故障级成因同拍置故障标志 / the fault flag paired with the cause
        _bFault := TRUE; _ePhase := E_DL_PraPhase.eFault; // 置锁存并迁故障相 / latch and migrate to the fault phase
    END_IF
E_DL_PraPhase.eSettle: // 稳定相：退出条件二（稳定窗到期 ｜ 使能丢失）
    IF NOT bEnable THEN // 使能丢失 / the enable was lost
        _ePhase := E_DL_PraPhase.eIdle; // 退回空闲 / back to idle
    ELSIF tonSettle.Q THEN // 稳定窗到期（拍 N 进入：本相起点 ｜ 本拍行为：拒绝新步进 ｜ 拍 N+1 转出：复评）
        _ePhase := E_DL_PraPhase.eEval; // 回评估相复评误差 / back to evaluate
    END_IF
E_DL_PraPhase.eDone: // 完成相：退出条件二（启动沿消失 ｜ 使能丢失），完成位由新循环起点清零
    IF (NOT bStart) OR (NOT bEnable) THEN // 启动电平消失或失能 / the start level dropped or the enable was lost
        _ePhase := E_DL_PraPhase.eIdle; // 回空闲相等下一轮 / back to idle for the next round
    END_IF
E_DL_PraPhase.eFault: // 故障相：成因锁存回放，唯一解除路径为 bReset 上升沿（R188）
    IF NOT bEnable THEN // 失能 / disabled
        _ePhase := E_DL_PraPhase.eIdle; // 迁空闲（锁存位仍须复位沿解除）/ migrate to idle, the latch still needs the reset edge
    END_IF
ELSE // 非法相位兜底（R6 / R128）/ the illegal phase fallback
    _eCause := E_DL_PraCause.ePhaseBad; _iErrLch := 105; // 故障级成因与码位：非法相位 / fault cause and code, an illegal phase
    bError := TRUE; // R45 配对：故障级成因同拍置故障标志 / the fault flag paired with the cause
    _bFault := TRUE; _ePhase := E_DL_PraPhase.eFault; // 置锁存并迁故障相 / latch and migrate to the fault phase
END_CASE
IF _bFault AND (_ePhase <> E_DL_PraPhase.eFault) THEN // 段尾迁移闸：任何锁存路径不得留在业务相（FB50-1④）
    _ePhase := E_DL_PraPhase.eFault; // 统一迁故障相 / force the fault phase
END_IF
// 段 8｜统一出口：命令、状态与码位单点映射（故障期命令保持末值，不再推进）
fVernierOut := _fVernAcc; // 色标偏移命令单点映射 / single point mapping of the offset command
fPhaseOut := _fPhaseA; // 版辊相位命令单点映射 / single point mapping of the phase command
fTensionOut := _fTensAcc; // 张力命令单点映射 / single point mapping of the tension command
nStepUsed := _nStep; // 步数单点映射 / single point mapping of the step count
nLadderIdx := _nLadder; // 阶梯编号单点映射 / single point mapping of the ladder index
bInTol := _bInTol; // 容差判据单点映射 / single point mapping of the tolerance verdict
bStepActive := (_ePhase = E_DL_PraPhase.eVern) OR (_ePhase = E_DL_PraPhase.eTens); // 等回执判据 / the waiting acknowledgement verdict
bBusy := bEnable AND (_ePhase <> E_DL_PraPhase.eIdle) AND (_ePhase <> E_DL_PraPhase.eDone) AND (_ePhase <> E_DL_PraPhase.eFault); // 运行位排除空闲完成与故障三相 / the busy bit excludes idle, done and fault
bDone := _bDone; // 完成位单点映射（保持式）/ single point mapping of the held done bit
bFault := _bFault; // 故障锁存单点映射 / single point mapping of the latch
IF _bFault THEN // 故障期回放锁存码，不在故障相按当下输入重推（R152）/ replay the latched code
    iErrCode := _iErrLch; // 锁存码回放 / replay the latched code
    bError := TRUE; // 故障标志与锁存位同源 / the fault flag shares the latch source
ELSE // 非故障期 / outside fault
    iErrCode := 0; // 无故障码 / no error code
    bError := FALSE; // 无故障标志 / no fault flag
END_IF
ePhase := _ePhase; // 相位出口单点映射 / single point mapping of the phase
END_FUNCTION_BLOCK

(* ---- FB_DL_PumpAlternationLead.st ---- *)
(*
    FB_DL_PumpAlternationLead —— 多泵轮换主备（小时均衡选主 + 故障切备锁存）
    ------------------------------------------------------------------
    组件名称  : FB_DL_PumpAlternationLead
    分类      : DL_Process / PumpGroup
    前缀      : FB_DL_
    版本      : 1.0.0
    溯源      : 借鉴点 —— 泵组轮换的通行工程语义：按累计运行小时选「最闲泵」作主泵、
                轮换周期到期强制换泵、在役泵故障时立即切备且故障泵被排除出候选集
                直至人工复位。该语义在公开工控资料中属常识性做法。
                clean-room 声明 —— 零代码行复制；选主算法、锁存结构、码位与双语文档
                全部本件自有，仅使用 IEC 61131-3 标准库 TON / R_TRIG。
                许可证 —— 本件 MIT；来源标签 self-std（道莅自有内规族），
                无第三方源码继承。
    平台      : 纯 IEC 61131-3，CODESYS 3.5 / TwinCAT 3 / InoProShop / Machine Expert 通用
    作者      : 道莅代码库 · PLC编程专家（R70 构建轮 · 批 2 · N5）
    ------------------------------------------------------------------
    功能说明  : 泵组固定 DL_PMP_N 台（默认 4 台，常数可改，全文件唯一定义）。
                选主规则：在所有「未被锁存排除」的泵中取累计运行小时最小者；
                小时完全相等的比较采用容差口径（不用浮点直比），相等时取小编号，
                故选主结果唯一、可复现。
                轮换规则：_tonRotate 以自复位口径产生周期脉冲（IN := bEn AND NOT Q，
                R188 禁靠外部沿清零）；脉冲拍强制排除当前主泵再选，实现主备交换。
                故障规则：abFault 为实时引脚输入，逐拍并入**每泵锁存位**
                _abFaultLatch，一旦置位即把该泵永久排除出候选集（本次运行期间），
                唯一解除边为 bReset 上升沿（R188 可到达的清除边）。
                锁存副本与实时镜像严格分离（历史教训 4）：判据只用 _abFaultLatch，
                abFault 引脚只用于「并入锁存」，二者绝不混用同一判据。
                小时累计：本件不自带计时基准，由上层按实际任务周期折算小时数后
                经 fScanHours 喂入（纯 IEC 口径，不依赖厂商 RTC 或 TIME 转换扩展），
                累计结果经 afRunHoursOut 出口回写上层保持区。
    错误码    : 16#0002_0201 组态非法（轮换周期 <= 0 或 fScanHours 非法），回放锁存 —— 故障级
                16#0002_0202 运行小时数组元素非法（负值 / 非有限），回放锁存 —— 故障级
                16#0002_0203 无可用泵（全部被锁存排除），输出全清零 —— 故障级
                16#0002_0204 主泵索引越界（内部一致性兜底，防数组越界访问）—— 故障级
    码位总账  : 0201 / 0202 / 0203 / 0204 用（均故障级）；无信息级码（本件不产生可观测的
                信息级事件，故不设，避免「声明了却永不赋值」）
    状态机    : N/A —— 无顺序相（选主为逐拍组合逻辑，轮换由定时脉冲驱动）；
                无 ENUM / CASE 可写，故无 CASE ELSE 兜底面
    边界与披露: 一 数组下标安全：全部 FOR 循环以常量 DL_PMP_N 为上下界（编译期确定），
                   另对 _nLead 做 1..N 显式校验并在越界时置 0204 且不索引数组，
                   两道防线同时存在，绝不出现下标越界读；
                二 组态闸（R272 逐项点名）：tRotate > T#0S；fScanHours 非有限闸 +
                   负值拦截；arRunHours 全元素非有限闸 + 负值拦截（累计小时不得为负）；
                三 加数饱和：小时累计结果按工程极限 DL_PMP_HCAP（1.0E12 h）夹住，
                   夹住后仍落在 LREAL 可表域内，故按「防御性夹住、不发码」处置 ——
                   该值在工程上不可达（1.0E12 h 远超设备寿命），发码只会产生
                   永不触发的死码位，违反「加码前须有现有输出组合不可观测的反证句」；
                四 失能（bEn = FALSE）：abCmd 全清零、bBusy 清零、轮换计时复位，
                   但每泵锁存位与小时累计**均不被清除**（失能非复位），须 bReset 解除；
                五 定时器 _tonRotate、沿实例 _rtReset 每周期无条件调用（规则 ⑦）；
                六 零全局变量、零 VAR_EXTERNAL、零物理地址、无除法。
    修订记录  : 2026-11-22 v1.0.0 首次入库（R70 构建轮 · 批 2 · N5）
*)
FUNCTION_BLOCK FB_DL_PumpAlternationLead
VAR_INPUT
    bEn         : BOOL := TRUE;                          (* 使能，[标志] / the enable *)
    bRunReq     : BOOL := FALSE;                          (* 泵组运行需求，[标志] / the group run request *)
    bReset      : BOOL := FALSE;                          (* 复位（上升沿解除故障锁存并清小时），[标志] / the reset, rising edge *)
    fScanHours  : LREAL := 0.0;                           (* 本周期折算小时数，[h]，由上层按任务周期喂入 / hours elapsed this scan *)
    arRunHours  : ARRAY[1..4] OF LREAL;                   (* 各泵累计运行小时（输入镜像），[h] / the per pump run hours, input image *)
    abFault     : ARRAY[1..4] OF BOOL;                    (* 各泵故障实时引脚，[标志] / the per pump live fault pins *)
    tRotate     : TIME := T#24H;                          (* 轮换周期，[ms]，须 > T#0S / the rotation period *)
END_VAR
VAR_OUTPUT
    nLead        : INT;                                   (* 当前主泵编号，0 = 无可用泵，[号] / the current lead pump number *)
    abCmd        : ARRAY[1..4] OF BOOL;                   (* 各泵运行命令出口，[标志] / the per pump run command *)
    afRunHoursOut : ARRAY[1..4] OF LREAL;                 (* 累计小时出口（上层回写保持区），[h] / the accumulated hours outlet *)
    bLeadChanged : BOOL;                                  (* 主泵切换单拍脉冲，[标志] / the lead change single scan pulse *)
    bBusy        : BOOL;                                  (* 轮换周期计时进行中，[标志] / the rotation period is timing *)
    bValid       : BOOL;                                  (* 出口可信（无锁存故障），[标志] / the outlets are trustworthy *)
    bError       : BOOL;                                  (* 故障标志，锁存故障时为 TRUE / the fault flag, raised while latched *)
    nErrCode     : UDINT;                                 (* 错误码，0 = 正常，锁存回放 / the error id, 0 = ok, replayed *)
END_VAR
VAR
    _rtReset       : R_TRIG;                              (* 复位上升沿实例（无条件调用）/ the reset rising edge instance *)
    _tonRotate     : TON;                                 (* 轮换周期计时实例（无条件调用，自复位口径）/ the rotation timer *)
    _abFaultLatch  : ARRAY[1..4] OF BOOL;                 (* 各泵故障锁存位，仅 bReset 解除 / the per pump latched fault *)
    _afHours       : ARRAY[1..4] OF LREAL;                (* 各泵小时工作副本（累计后出口），[h] / the per pump working copy *)
    _nLead         : INT;                                 (* 当前主泵寄存器，[号] / the lead pump register *)
    _nPrevLead     : INT;                                 (* 上拍主泵快照（切换沿基准），[号] / the previous lead snapshot *)
    _bFault        : BOOL;                                (* 块级故障锁存位 / the block level fault latch *)
    _nCodeLatch    : UDINT;                               (* 锁存成因码，故障期回放 / the latched cause code *)
    _bCfgBad       : BOOL;                                (* 组态非法标志（逐拍重算）/ the configuration fault flag *)
    _bHoursBad     : BOOL;                                (* 小时数组非法标志（逐拍重算）/ the hour array fault flag *)
    _bRun          : BOOL;                                (* 运行许可 = 使能 且 无锁存故障 / the run permit *)
    _bRotNeed      : BOOL;                                (* 本拍需强制轮换（定时脉冲）/ the rotation is due this scan *)
    _i             : INT;                                 (* 循环下标，[号] / the loop index *)
    _nBest         : INT;                                 (* 本轮选出的候选泵号，0 = 无，[号] / the selected candidate *)
    _nIdx          : INT;                                 (* 已校验的下标副本（索引前必判），[号] / the validated index copy *)
    _fBest         : LREAL;                               (* 候选最小小时值，[h] / the smallest hours found *)
    _bConsider     : BOOL;                                (* 该泵是否进入本轮候选，[标志] / whether the pump is a candidate *)
    _bTie          : BOOL;                                (* 小时相等（容差内）判据结果，[标志] / the tie verdict *)
END_VAR
VAR CONSTANT
    DL_PMP_N       : INT := 4;                            (* 泵台数（与数组声明同源），[台] / the pump count, matching the arrays *)
    DL_PMP_FMAX    : LREAL := 1.0E30;                     (* 非有限筛查幅值上限，[h] / the finiteness screening cap *)
    DL_PMP_HTOL    : LREAL := 1.0E-9;                     (* 小时相等比较容差，[h] / the hours equality tolerance *)
    DL_PMP_HCAP    : LREAL := 1.0E12;                     (* 小时累计上限（工程极限，夹住），[h] / the hours accumulation cap *)
    DL_PMP_NONE    : INT := 0;                            (* 无可用泵的哨兵值，[号] / the no-available-pump sentinel *)
END_VAR

// 段 1｜出口预置（R256 统一出口预置）/ segment 1, preset every outlet
bLeadChanged := FALSE;                     // 切换脉冲预清零 / preset the change pulse false
bBusy        := FALSE;                     // 忙碌标志预清零 / preset the busy flag false
bValid       := FALSE;                     // 可用标志预置假，健康路径再置真 / preset valid false, set in the healthy path
bError       := FALSE;                     // 故障标志预清零 / preset the error flag false
nErrCode     := 0;                         // 错误码预置无错 / preset the code to zero
_bRotNeed    := FALSE;                     // 轮换需求预清零 / preset the rotation need false
FOR _i := 1 TO DL_PMP_N DO                 // 常量上下界，下标安全 / constant bounds, indices safe
    abCmd[_i] := FALSE;                    // 各泵命令预清零（失能安全方向）/ preset every command off
    afRunHoursOut[_i] := _afHours[_i];     // 小时出口镜像工作副本 / mirror the working copy
END_FOR

// 段 2｜沿实例与定时器无条件调用（规则 ⑦）/ segment 2, the edge instance and the timer, called unconditionally
_rtReset(CLK := bReset);                               // 复位沿，每周期无条件刷新 / the reset edge, refreshed every scan
_tonRotate(IN := (bEn AND NOT _tonRotate.Q), PT := tRotate); // 轮换周期自复位计时（R188）/ the self resetting rotation timer

// 段 3｜复位解除：唯一可到达的清除边（R188）/ segment 3, the only reachable clearing edge
IF _rtReset.Q THEN                         // 复位上升沿 / the reset rising edge
    _bFault     := FALSE;                  // 解除块级故障锁存 / release the block fault latch
    _nCodeLatch := 0;                      // 清锁存码 / clear the latched code
    FOR _i := 1 TO DL_PMP_N DO             // 常量上下界 / constant bounds
        _abFaultLatch[_i] := FALSE;        // 解除各泵故障锁存 / release every per pump latch
    END_FOR
END_IF

// 段 4｜组态闸：轮换周期与扫描小时数（R272 逐项点名）/ segment 4, the configuration gate
_bCfgBad := (tRotate <= T#0S)                                     // 轮换周期非正 / a non positive rotation period
         OR (fScanHours < 0.0)                                    // 扫描时长为负 / a negative elapsed time
         OR (fScanHours <> fScanHours) OR ((fScanHours - fScanHours) <> 0.0) OR (ABS(fScanHours) > DL_PMP_FMAX);

// 段 5｜小时数组闸：全元素非有限 + 负值拦截 / segment 5, the hour array gate
_bHoursBad := FALSE;                       // 逐拍重算 / recomputed every scan
FOR _i := 1 TO DL_PMP_N DO                 // 常量上下界 / constant bounds
    IF (arRunHours[_i] <> arRunHours[_i]) OR ((arRunHours[_i] - arRunHours[_i]) <> 0.0)
       OR (ABS(arRunHours[_i]) > DL_PMP_FMAX) OR (arRunHours[_i] < 0.0) THEN // 元素非法 / an illegal element
        _bHoursBad := TRUE;                // 标记非法 / flag it
    END_IF
END_FOR

// 段 6｜首次成因锁存（故障期不重推断，R189）/ segment 6, the first cause latch
IF NOT _bFault THEN                        // 未锁存才登记 / register only while healthy
    IF _bCfgBad THEN                       // 组态非法优先 / the configuration first
        _bFault     := TRUE;               // 置锁存 / latch it
        _nCodeLatch := 16#0002_0201;       // 故障级：组态非法 / fault level: an illegal configuration
    ELSIF _bHoursBad THEN                  // 小时数组非法 / the hour array is illegal
        _bFault     := TRUE;               // 置锁存 / latch it
        _nCodeLatch := 16#0002_0202;       // 故障级：小时数组非法 / fault level: the hour array is illegal
    END_IF
END_IF

// 段 7｜实时故障引脚并入每泵锁存位（锁存副本与实时镜像分离，历史教训 4）/ segment 7, merge the live pins into the latches
FOR _i := 1 TO DL_PMP_N DO                 // 常量上下界 / constant bounds
    IF abFault[_i] THEN                    // 实时引脚为真 / the live pin is true
        _abFaultLatch[_i] := TRUE;         // 并入锁存（只增不减，唯一解除边见段 3）/ merge into the latch, released only in segment 3
    END_IF
END_FOR

// 段 8｜运行许可与轮换需求 / segment 8, the run permit and the rotation request
_bRun     := bEn AND NOT _bFault;          // 使能且无锁存故障 / enabled and not latched
_bRotNeed := _bRun AND bRunReq AND _tonRotate.Q; // 周期到且确有运行需求才轮换 / rotate when due and actually demanded
bBusy     := _bRun AND bRunReq AND NOT _tonRotate.Q; // 轮换周期计时中 / the rotation period is timing

// 段 9｜小时累计（仅对当前在役主泵累加）与出口 / segment 9, accumulate the hours of the running lead
IF _bRun THEN                              // 运行许可成立 / the run permit holds
    FOR _i := 1 TO DL_PMP_N DO             // 常量上下界 / constant bounds
        _afHours[_i] := arRunHours[_i];    // 先取输入镜像 / take the input image first
    END_FOR
    IF bRunReq THEN                        // 确有运行需求时主泵才计小时 / only a demanded lead accumulates
        _nIdx := _nLead;                   // 取待校验下标 / take the index to validate
        IF (_nIdx >= 1) AND (_nIdx <= DL_PMP_N) THEN   // 索引先判（防越界，规则 ④）/ validate before indexing
            _afHours[_nIdx] := _afHours[_nIdx] + fScanHours;   // 累加本周期小时 / add the elapsed hours
            IF _afHours[_nIdx] > DL_PMP_HCAP THEN              // 超工程极限 / beyond the engineering cap
                _afHours[_nIdx] := DL_PMP_HCAP;                // 夹住（夹住仍在实数可表域内）/ clamp it
            END_IF
        END_IF
    END_IF
    FOR _i := 1 TO DL_PMP_N DO             // 常量上下界 / constant bounds
        afRunHoursOut[_i] := _afHours[_i]; // 小时出口回写 / write the hours outlet
    END_FOR
ELSE                                       // 失能或锁存故障 / disabled or latched
    FOR _i := 1 TO DL_PMP_N DO             // 常量上下界 / constant bounds
        _afHours[_i] := arRunHours[_i];    // 工作副本照旧镜像（不做累计）/ mirror without accumulation
        afRunHoursOut[_i] := _afHours[_i]; // 出口照旧（小时不被失能清零）/ the outlet is not cleared by a disable
    END_FOR
END_IF

// 段 10｜选主：最闲泵，轮换拍排除当前主泵 / segment 10, the lead selection
_nPrevLead := _nLead;                      // 上拍主泵快照（切换沿基准）/ snapshot the previous lead
_nBest     := DL_PMP_NONE;                 // 候选初值：无 / the candidate starts empty
_fBest     := DL_PMP_FMAX;                 // 最小小时初值为筛查上界 / the smallest hours starts at the cap
IF _bRun THEN                              // 运行许可成立 / the run permit holds
    FOR _i := 1 TO DL_PMP_N DO             // 常量上下界 / constant bounds
        _bConsider := NOT _abFaultLatch[_i];                            // 未被锁存排除 / not excluded by the latch
        IF _bRotNeed AND (_i = _nLead) THEN                             // 轮换拍排除当前主泵 / exclude the current lead on a rotation
            _bConsider := FALSE;                                        // 退出候选 / drop it from the candidates
        END_IF
        IF _bConsider THEN                                              // 候选泵 / a candidate
            _bTie := ABS(_afHours[_i] - _fBest) <= DL_PMP_HTOL;         // 小时相等（容差口径）/ an hours tie within tolerance
            IF (_fBest > (DL_PMP_FMAX - DL_PMP_HTOL)) OR (_afHours[_i] < _fBest) OR _bTie THEN
                IF NOT ((_nBest <> DL_PMP_NONE) AND _bTie) THEN          // 已有候选且相等时保留小编号 / keep the lower number on a tie
                    _fBest := _afHours[_i];                             // 刷新最小值 / refresh the minimum
                    _nBest := _i;                                       // 记录候选泵号 / record the candidate
                END_IF
            END_IF
        END_IF
    END_FOR
    IF _nBest = DL_PMP_NONE THEN                                   // 轮换拍把唯一可用泵排除了 / the rotation excluded the only pump
        _nIdx := _nLead;                                           // 取待校验下标 / take the index to validate
        IF (_nIdx >= 1) AND (_nIdx <= DL_PMP_N) THEN               // 索引先判 / validate first
            IF NOT _abFaultLatch[_nIdx] THEN                       // 原主泵仍健康 / the previous lead is still healthy
                _nBest := _nIdx;                                   // 回落保持原主泵 / fall back to the previous lead
            END_IF
        END_IF
    END_IF
    IF _nBest = DL_PMP_NONE THEN                                   // 确实无可用泵 / truly no pump available
        _bFault     := TRUE;                                       // 锁存故障 / latch the fault
        _nCodeLatch := 16#0002_0203;                               // 故障级：无可用泵 / fault level: no pump available
    END_IF
END_IF

// 段 11｜主泵索引校验与命令出口（名实双出口同源，R191）/ segment 11, validate the lead and drive the outlets
IF _bRun AND NOT _bFault THEN              // 健康运行 / healthy and running
    _nIdx := _nBest;                       // 取待校验下标 / take the index to validate
    IF (_nIdx >= 1) AND (_nIdx <= DL_PMP_N) THEN   // 索引先判（规则 ④）/ validate before indexing
        _nLead := _nIdx;                   // 提交主泵寄存器 / commit the lead register
        IF bRunReq THEN                    // 有运行需求 / a run is demanded
            abCmd[_nIdx] := TRUE;          // 仅主泵运行（单泵运行策略）/ only the lead runs
        END_IF
        bValid := TRUE;                    // 出口可信 / the outlets are trustworthy
    ELSE                                   // 内部一致性失败 / an internal consistency failure
        _nLead      := DL_PMP_NONE;        // 主泵清为无 / clear the lead
        _bFault     := TRUE;               // 锁存故障 / latch the fault
        _nCodeLatch := 16#0002_0204;       // 故障级：主泵索引越界 / fault level: the lead index out of range
    END_IF
END_IF

// 段 12｜出口映射（单点写入，无自赋值）/ segment 12, the outlet mapping
nLead        := _nLead;                    // 主泵号出口 / the lead number outlet
bLeadChanged := (_nLead <> _nPrevLead);    // 主泵切换单拍脉冲（整数直比，无浮点面）/ the lead change pulse
bError       := _bFault;                   // 名实双出口：故障位与锁存同源（R191）/ both outlets share the latch
nErrCode     := _nCodeLatch;               // 锁存码回放 / replay the latched code
IF _bFault THEN                            // 锁存故障相 / the latched fault phase
    bValid := FALSE;                       // 出口不可信 / the outlets are not trustworthy
    FOR _i := 1 TO DL_PMP_N DO             // 常量上下界 / constant bounds
        abCmd[_i] := FALSE;                // 全泵命令清零（失效安全）/ all commands off
    END_FOR
END_IF
END_FUNCTION_BLOCK

(* ---- FB_DL_PumpChangeoverSeq.st ---- *)
(*==============================================================================
 * 组件名称 (Component)  : FB_DL_PumpChangeoverSeq
 * 所属子库 (Sublibrary) : DL_Process
 * 当前版本 (Version)    : 1.0.0
 * 兼容性 (Platform)     : CODESYS 3.5 / TwinCAT 3 / 汇川 InoProShop / Machine Expert
 *                         仅依赖纯 IEC 61131-3 标准元素，零厂商方言
 * 功能描述 (Function)   : 冷冻/冷却水泵加减机：供回水温差与目标温差比较，死区
 *                         ±0.5 摄氏度内保持；滞消频宽后折算级数需求（下限 1，
 *                         水泵不保备机——与风机阵列的差异点）；每 tick 至多切换
 *                         1 台，tMinRun/tMinStop 闸门防频繁启停；轮值按运行小时
 *                         均衡选台。温差传感器无效 → 保持当前组合只报码不切换。
 * 溯源 (Origin)         : 道莅 clean-room 防御性实现
 * 本文件内含 (Contains) : TYPE E_DL_ChgoverErr / FUNCTION_BLOCK FB_DL_PumpChangeoverSeq
 * 依赖 (Depends)        : 无 DL_ 内部依赖；Standard.library TON 实例
 * 红线自检 (Redline)    : 无外部全局变量、无硬件地址直引 ｜ 全变量中英双语同行注释
 *                         数组下界常量提取 + 级数钳位 [1,N] + 非有限温差不切换 ｜
 *                         枚举成员全部显式赋值 ｜ TON 实例每周期无条件调用 ｜
 *                         CASE 含 ELSE 兜底 ｜ 与风机阵列共纪律但零共享实例
 * 错误码表 (Codes)      : 16#0005_0426 就绪
 *                         16#0005_0427 信息级 温差在死区（保持，含传感器无效保持）
 *                         16#0005_0428 信息级 加机中
 *                         16#0005_0429 信息级 减机中
 *                         16#0005_042A 信息级 闸门等待（最短时序未满足）
 * 修订历史 (Revision)   : 2026-11-17  v1.0.0  首版入库 · R27 · 阶段三批 4
 * 验收向量 (Acceptance) : 目标 5 摄氏度，实测 7.0 → 需求加 1 台并 0428；
 *                         实测 6.0（死区内）→ 保持 0427；切换后 tMinRun 内再要
 *                         切换 → 042A 只记不切
 *============================================================================*)

(*-----------------------------------------------------------------------------
 * 枚举: E_DL_ChgoverErr（归属 DL_Process，与 FB_DL_PumpChangeoverSeq 同文件）
 *----------------------------------------------------------------------------*)
TYPE E_DL_ChgoverErr :
(
    eReady   := 16#0005_0426,   // 就绪 / Ready
    eDeadband:= 16#0005_0427,   // 信息级：温差在死区或传感器无效（保持）/ Info: deadband or invalid sensor, hold
    eAddRun  := 16#0005_0428,   // 信息级：加机中 / Info: adding a pump
    eSubRun  := 16#0005_0429,   // 信息级：减机中 / Info: shedding a pump
    eGateWait:= 16#0005_042A    // 信息级：闸门等待 / Info: minimum-timing gate waiting
);
END_TYPE

(*==============================================================================
 * 功能块: FB_DL_PumpChangeoverSeq
 * 调用约定: 每个扫描周期无条件调用一次；aNRunHrs 由调用方按索引注入。
 *============================================================================*)
FUNCTION_BLOCK FB_DL_PumpChangeoverSeq
VAR_INPUT
    fDeltaT_C    : REAL;                     // 供回水温差 [摄氏度] / Supply-return temperature difference [degC]
    fDeltaTSet_C : REAL := 5.0;              // 目标温差 [摄氏度]，默认 5 / Target temperature difference [degC]
    aNRunHrs     : ARRAY[1..6] OF UDINT;     // 各泵累计运行小时 [小时] / Run hours per pump [h]
    uPumpTotal   : UINT := 6;                // 装机泵数 [台]，有效域 1~6 / Installed pump count [pumps]
    tMinRun      : TIME := T#60S;            // 最短运行时长 [秒] / Minimum run time [s]
    tMinStop     : TIME := T#60S;            // 最短停机时长 [秒] / Minimum stop time [s]
END_VAR
VAR_OUTPUT
    auPumpCmd    : ARRAY[1..6] OF BOOL;      // 各泵启停指令 / Pump start/stop commands
    uRunCount    : UINT;                     // 实际运行泵数 [台] / Actual running pump count [pumps]
    eErr         : E_DL_ChgoverErr;          // 错误码 / Error code
END_VAR
VAR
    tonGateRun   : TON;                      // 最短运行闸门定时器（无条件调用）/ Min-run gate timer
    tonGateStop  : TON;                      // 最短停机闸门定时器（无条件调用）/ Min-stop gate timer
    bGateArmed   : BOOL;                     // 闸门武装标志（切换后置位）/ Gate armed flag
    bSwitchCycle : BOOL;                     // 本拍为切换拍（定时器 IN 强制断流）/ Switch-scan flag, forces timer reset
    fSetUse      : REAL;                     // 生效目标温差 [摄氏度] / Effective target difference [degC]
    fDev_C       : REAL;                     // 温差偏差 [摄氏度] / Temperature difference deviation [degC]
    uTotalUse    : UINT;                     // 生效泵数（钳位后）[台] / Effective pump count [pumps]
    uStageNeed   : UINT;                     // 级数需求 [台] / Stage demand [pumps]
    uIdxBest     : UINT;                     // 候选切换泵索引 [台序] / Candidate pump index
    nPickHrs     : UDINT;                    // 候选比较基准小时 [小时] / Candidate comparison baseline [h]
    i            : INT;                      // 数组循环索引 / Array loop index
    bSensorOk    : BOOL;                     // 温差传感器有效判据 / Temperature sensor validity predicate
    bInit        : BOOL;                     // 首扫初始化标志 / First-scan init flag
END_VAR
VAR CONSTANT
    DL_CHG_IDX_MAX   : INT  := 6;            // 阵列容量上限（数组下界常量提取）/ Array capacity upper bound
    DL_CHG_TOTAL_MAX : UINT := 6;            // 装机泵数上限 [台] / Installed count upper bound [pumps]
    DL_CHG_STAGE_MIN : UINT := 1;            // 级数下限 1 台（水泵不保备机，与风机阵列差异）/ Stage lower bound, one pump minimum
    DL_CHG_DEADBAND  : REAL := 0.5;          // 死区半宽 [摄氏度] / Deadband half width [degC]
    DL_CHG_STAGE_C   : REAL := 2.0;          // 级数折算温差步长 [摄氏度每台] / Stage temperature step [degC per pump]
    DL_CHG_INF_MAX   : REAL := 1.0E30;       // 非有限值判定幅值上限 / Magnitude bound for finite-value check
    DL_CHG_ZERO      : REAL := 0.0;          // 零值常量，避免裸字面量 / Zero constant
END_VAR

(*------------------------------------------------------------------------------
 * 段 1｜TON 实例每周期无条件调用（仅 IN 条件化）：切换拍强制断流以复位计时
 *----------------------------------------------------------------------------*)
tonGateRun(IN := bGateArmed AND NOT bSwitchCycle, PT := tMinRun);     // 运行闸计时 / min-run gate timing
tonGateStop(IN := bGateArmed AND NOT bSwitchCycle, PT := tMinStop);   // 停机闸计时 / min-stop gate timing

(*------------------------------------------------------------------------------
 * 段 2｜首扫初始化：指令数组全停
 *----------------------------------------------------------------------------*)
IF NOT bInit THEN
    FOR i := 1 TO DL_CHG_IDX_MAX DO
        auPumpCmd[i] := FALSE;                           // 默认全停 / default all stopped
    END_FOR
    bInit := TRUE;                                       // 首扫完成 / first scan done
END_IF

(*------------------------------------------------------------------------------
 * 段 3｜泵数钳位与目标温差兜底
 *----------------------------------------------------------------------------*)
uTotalUse := uPumpTotal;                                 // 泵数工作副本 / total working copy
IF uTotalUse > DL_CHG_TOTAL_MAX THEN
    uTotalUse := DL_CHG_TOTAL_MAX;                       // 泵数上限钳位 / total capped
ELSIF uTotalUse < DL_CHG_STAGE_MIN THEN
    uTotalUse := DL_CHG_STAGE_MIN;                       // 泵数下限钳位 / total floored
END_IF
fSetUse := fDeltaTSet_C;                                 // 目标工作副本 / target working copy
IF (fSetUse <> fSetUse) OR (fSetUse <= DL_CHG_ZERO) OR (fSetUse > DL_CHG_INF_MAX) THEN
    fSetUse := 5.0;                                      // 目标非法按 5 摄氏度兜底 / illegal target falls back to 5 degC
END_IF

(*------------------------------------------------------------------------------
 * 段 4｜传感器有效性与偏差计算：无效则保持当前组合只报码
 *----------------------------------------------------------------------------*)
bSensorOk := (fDeltaT_C = fDeltaT_C) AND (ABS(fDeltaT_C) <= DL_CHG_INF_MAX) AND (fDeltaT_C >= DL_CHG_ZERO);   // 温差有效 / difference validity
eErr := E_DL_ChgoverErr.eReady;                          // 预置就绪 / preset ready
uStageNeed := uRunCount;                                 // 需求缺省 = 当前运行数（保持）/ demand defaults to current count
IF NOT bSensorOk THEN
    eErr := E_DL_ChgoverErr.eDeadband;                   // 信息级：传感器无效保持（与死区共用，反证句：均为不切换）/ info: invalid sensor, hold
ELSE
    fDev_C := fDeltaT_C - fSetUse;                       // 温差偏差 [摄氏度] / difference deviation [degC]
    IF (fDev_C > -DL_CHG_DEADBAND) AND (fDev_C < DL_CHG_DEADBAND) THEN
        eErr := E_DL_ChgoverErr.eDeadband;               // 信息级：死区内保持 / info: inside deadband, hold
    ELSIF fDev_C > DL_CHG_ZERO THEN
        // 温差偏高：需要加机（级数需求按偏差折算，上限泵数）/ positive deviation: more pumps
        uStageNeed := uRunCount + UDINT_TO_UINT(REAL_TO_UDINT(ROUND(fDev_C / DL_CHG_STAGE_C)));   // 需求级数折算 [台] / stage demand
        IF uStageNeed <= uRunCount THEN
            uStageNeed := uRunCount + 1;                 // 至少加 1 台（ROUND 归零时保底）/ at least one more pump
        END_IF
        IF uStageNeed > uTotalUse THEN
            uStageNeed := uTotalUse;                     // 需求上限钳位（不保备机）/ demand capped at total
        END_IF
    ELSE
        // 温差偏低：需要减机（下限 1 台）/ negative deviation: fewer pumps, one minimum
        IF fDev_C < -DL_CHG_STAGE_C THEN
            uStageNeed := uRunCount - 1;                 // 偏差超一个步长：减 1 台 / shed one pump
        ELSE
            uStageNeed := uRunCount;                     // 偏差未超步长：保持 / hold, within one step
        END_IF
        IF uStageNeed < DL_CHG_STAGE_MIN THEN
            uStageNeed := DL_CHG_STAGE_MIN;              // 下限钳位 1 台 / floored at one pump
        END_IF
    END_IF
END_IF

(*------------------------------------------------------------------------------
 * 段 5｜每 tick 至多切换 1 台：加机选小时最少，减机选小时最多
 *----------------------------------------------------------------------------*)
uIdxBest := 0;                                           // 候选索引清零（0 = 无候选）/ candidate reset
nPickHrs := 0;                                           // 基准清零 / baseline reset
IF uRunCount > uStageNeed THEN
    IF bGateArmed AND NOT tonGateRun.Q THEN
        eErr := E_DL_ChgoverErr.eGateWait;               // 信息级：闸门等待（只记不切）/ info: gate waiting
    ELSE
        nPickHrs := 0;                                   // 最多小时基准从 0 起比 / max search baseline
        FOR i := 1 TO UINT_TO_INT(uTotalUse) DO
            IF auPumpCmd[i] THEN
                IF (uIdxBest = 0) OR (aNRunHrs[i] >= nPickHrs) THEN
                    uIdxBest := INT_TO_UINT(i);          // 候选更新（运行最久）/ candidate updated
                    nPickHrs := aNRunHrs[i];             // 基准更新 / baseline updated
                END_IF
            END_IF
        END_FOR
        IF uIdxBest > 0 THEN
            eErr := E_DL_ChgoverErr.eSubRun;             // 信息级：减机中 / info: shedding
        END_IF
    END_IF
ELSIF uRunCount < uStageNeed THEN
    IF bGateArmed AND NOT tonGateStop.Q THEN
        eErr := E_DL_ChgoverErr.eGateWait;               // 信息级：闸门等待（只记不切）/ info: gate waiting
    ELSE
        nPickHrs := 16#FFFF_FFFF;                        // 最少小时基准从满值起比 / min search baseline
        FOR i := 1 TO UINT_TO_INT(uTotalUse) DO
            IF NOT auPumpCmd[i] THEN
                IF aNRunHrs[i] <= nPickHrs THEN
                    uIdxBest := INT_TO_UINT(i);          // 候选更新（停机最久近似小时最少）/ candidate updated
                    nPickHrs := aNRunHrs[i];             // 基准更新 / baseline updated
                END_IF
            END_IF
        END_FOR
        IF uIdxBest > 0 THEN
            eErr := E_DL_ChgoverErr.eAddRun;             // 信息级：加机中 / info: adding
        END_IF
    END_IF
END_IF

(*------------------------------------------------------------------------------
 * 段 6｜执行切换：切换拍置武装并强制定时器断流复位
 *----------------------------------------------------------------------------*)
bSwitchCycle := FALSE;                                   // 切换拍标志默认 FALSE / switch-scan flag defaults FALSE
IF uIdxBest > 0 THEN
    auPumpCmd[UINT_TO_INT(uIdxBest)] := NOT auPumpCmd[UINT_TO_INT(uIdxBest)];   // 执行切换 / execute the switch
    bGateArmed := TRUE;                                  // 闸门武装 / gate armed
    bSwitchCycle := TRUE;                                // 切换拍标志（下拍定时器重新计时）/ switch-scan flag
END_IF

(*------------------------------------------------------------------------------
 * 段 7｜运行泵数统计与容量外指令清扫（防越界残留）
 *----------------------------------------------------------------------------*)
uRunCount := 0;                                          // 运行泵数清零 / running count reset
FOR i := 1 TO DL_CHG_IDX_MAX DO
    IF i > UINT_TO_INT(uTotalUse) THEN
        auPumpCmd[i] := FALSE;                           // 容量外指令强制撤销 / force FALSE beyond capacity
    ELSIF auPumpCmd[i] THEN
        uRunCount := uRunCount + 1;                      // 运行泵数累加 [台] / running count incremented
    END_IF
END_FOR
END_FUNCTION_BLOCK

(* ---- FB_DL_PumpDownEnvelopeMonitor.st ---- *)
(*==============================================================================
 * 组件名称 (Component)  : FB_DL_PumpDownEnvelopeMonitor
 * 所属子库 (Sublibrary) : DL_Process
 * 当前版本 (Version)    : 1.0.1
 * 命名说明 (Naming)     : 本库已存在 FB_DL_ChamberPumpDownProfile（早期入库，引脚为包络上界
 *                         与停滞极差口径，码位 0005_01F2/01F3/0330~0332）。R28 计划书序 13
 *                         的引脚口径（seg1End/seg2End 段界 + 斜率包络 + 抽速早停建议）与之
 *                         不兼容，且同名会与已注册组件撞名，故按「段界斜率包络」语义另立
 *                         本名，旧件保持不动。命名归属待总监裁定。
 * 兼容性 (Platform)     : CODESYS 3.5 / TwinCAT 3 / 汇川 InoProShop（纯标准元素，零方言）
 * 功能描述 (Function)   : 抽气曲线三段包络监视与抽速早停建议。按段界压强把抽气过程分为
 *                         粗抽 / 过渡 / 精抽三段，逐段用采样斜率与最小抽速比较：低于包络只
 *                         给早停**建议**（bSlowWarn），绝不切泵；压强非有限立即停段并报故障；
 *                         段超时只建议不切断。不做泵启停、不做阀门时序、不做泄漏率诊断。
 *                         交付门槛：斜率用时间转换链换算秒，须在 CODESYS / TwinCAT /
 *                         InoProShop 三平台各编译验证一次。
 * 溯源 (Origin)         : 道莅 clean-room 防御性实现
 * 本文件内含 (Contains) : TYPE E_DL_PumpSeg / FUNCTION_BLOCK FB_DL_PumpDownEnvelopeMonitor
 * 依赖 (Depends)        : 无（仅 Standard.library 的 ABS / TIME_TO_LREAL）
 * 红线自检 (Redline)    : 无外部全局变量、无硬件地址直引 ｜ 全变量中英双语同行注释
 *                         最小抽速与采样周期判零防除零 ｜ 段界反置判组态错 ｜ 压强非有限即
 *                         停段（不可读不许推进段）｜ 采样与段超时定时器无条件周期刷新 ｜
 *                         枚举显式赋值 ｜ CASE 含 ELSE 兜底
 * 错误码表 (Codes)      : 16#0005_0435 就绪（各段正常或非抽气期）
 *                         16#0005_0436 预留：本版不发码（下一轮区间起点，禁止回填）
 *                         16#0005_0437 故障级 组态非法（段界反置或最小抽速 ≤0、采样周期出域）
 *                         16#0005_0438 信息级 段超时，只给早停建议（不切泵、不置故障级标志）
 *                         16#0005_0439 故障级 压强非有限，停段（uSeg=9，不可读不许推进段）
 * 修订历史 (Revision)   : 2026-11-17  v1.0.0  首版入库 · R28 · 阶段三批 3（因撞名另立名）
 *                         2026-11-17  v1.0.1  终审修复：①早停建议改为段内锁存派生输出，新循环
 *                                    起点同拍清零（原「置位后永不清」会向上位留幽灵建议）；
 *                                    ②故障码改由锁存码回放，原「守不住原码」会把组态故障错
 *                                    报成压强故障· R28 · 阶段四
 * 验收向量 (Acceptance) : 正向 101→10 kPa/30 s（3.03 kPa/s）+ 10→1 kPa/45 s（0.2 kPa/s）、
 *                         最小抽速 0.1 → 全程合格、bProfileOk
 *                         反向 段拖到 200 s（0.045 kPa/s 低于 0.1）→ bSlowWarn 且不置故障；
 *                         段界反置 → 16#0005_0437；压强给 NaN → uSeg=9 + 16#0005_0439
 *============================================================================*)

(*-----------------------------------------------------------------------------
 * 枚举: E_DL_PumpSeg（归属本功能块，同文件发布，全库唯一定义）
 *----------------------------------------------------------------------------*)
TYPE E_DL_PumpSeg :
(
    eIdle  := 0,    // 待机：泵未运行 / Idle, the pump is not running
    eRough := 1,    // 粗抽段：压强高于段界 1 / Rough segment above boundary one
    eTrans := 2,    // 过渡段：介于段界 1 与段界 2 / Transition between the two boundaries
    eFine  := 3,    // 精抽段：低于段界 2 / Fine segment below boundary two
    eDone  := 4,    // 完成：全程达标 / Done, the whole profile was acceptable
    eFault := 9     // 故障：读数不可信，停段 / Fault, the reading is untrustworthy and the segment stops
);
END_TYPE

FUNCTION_BLOCK FB_DL_PumpDownEnvelopeMonitor
VAR_INPUT
    bEnable       : BOOL := FALSE;        // 使能 / Enable
    bPumpOn       : BOOL := FALSE;        // 泵运行中 / Pump running
    fPress_kPa    : REAL := 101.3;        // 腔体压强 [kPa(abs)] / Chamber pressure in kilopascal absolute
    fSeg1End_kPa  : REAL := 10.0;         // 段界 1 压强 [kPa(abs)]，须 > 段界 2 / Boundary one, must exceed boundary two
    fSeg2End_kPa  : REAL := 1.0;          // 段界 2 压强 [kPa(abs)] / Boundary two
    fSlopeMin_kPas : REAL := 0.1;         // 各段最小抽速 [kPa/s]，域 0.001~10 / Minimum slope, domain 0.001 to 10
    tSampleTime   : TIME := T#100MS;      // 采样周期 [ms]，域 10~1000 / Sampling period, domain 10 to 1000 ms
    tSegMax       : TIME := T#1800S;      // 单段超时 [ms]，域 1~1800 s / Per-segment timeout
END_VAR
VAR_OUTPUT
    fSeg1Slope_kPas : REAL;               // 段 1 实测斜率 [kPa/s] / Measured slope of segment one
    fSeg2Slope_kPas : REAL;               // 段 2 实测斜率 [kPa/s] / Measured slope of segment two
    uSeg          : UINT;                 // 段号 0 待机 1 粗抽 2 过渡 3 精抽 4 完成 9 故障 [—] / Segment number
    bSlowWarn     : BOOL;                 // 低于包络（早停建议） / Below the envelope, early-stop advice
    bProfileOk    : BOOL;                 // 全程合格 / The whole profile is acceptable
    eErr          : UDINT;                // 错误码，段位 16#0005_xxxx / Error code in segment 16#0005_xxxx
END_VAR
VAR
    _eSeg         : E_DL_PumpSeg := E_DL_PumpSeg.eIdle; // 当前段 / Current segment
    _bInit        : BOOL := FALSE;        // 首扫标志，取非判定 / First-scan flag, tested negated
    _bCfgOk       : BOOL;                 // 组态合法标志 / Configuration valid flag
    _bHasSample   : BOOL := FALSE;        // 已有上一拍样本 / A previous sample exists
    _bSlowLatch   : BOOL := FALSE;        // 早停建议锁存（段内保持） / Early-stop advice latched inside a segment
    _uLatchCode   : UDINT;                // 故障锁存码载体（回放用） / Latch code carrier for the replay
    _bS1Judged    : BOOL := FALSE;        // 段 1 已判定标志 / Segment one already judged
    _bS2Judged    : BOOL := FALSE;        // 段 2 已判定标志 / Segment two already judged
    _fPrev_kPa    : REAL := 0.0;          // 上一拍压强 [kPa(abs)] / Previous pressure sample
    _fSampleSec   : REAL := 0.1;          // 采样周期换算秒 [s] / Sampling period in seconds
    _fSlope       : REAL;                 // 本拍斜率 [kPa/s] / Slope of this scan
    _rtrigSample  : R_TRIG;               // 采样节拍沿 / Sample tick edge
    _tonSample    : TON;                  // 采样周期计时（自复位） / Sampling period timer, self resetting
    _tonSeg       : TON;                  // 段超时计时 / Segment timeout timer
END_VAR
VAR CONSTANT
    DL_PD_READY    : UDINT := 16#0005_0435;  // 就绪码 / Ready code
    DL_PD_CFG_BAD  : UDINT := 16#0005_0437;  // 故障级组态非法码 / Fault code for bad configuration
    DL_PD_SEG_TO   : UDINT := 16#0005_0438;  // 信息级段超时码 / Info code for a segment timeout
    DL_PD_PRESS_BAD : UDINT := 16#0005_0439; // 故障级压强非有限码 / Fault code for a non-finite pressure
    DL_PD_SLOPE_LO : REAL := 0.001;          // 最小抽速下限 [kPa/s] / Minimum slope lower bound
    DL_PD_SLOPE_HI : REAL := 10.0;           // 最小抽速上限 [kPa/s] / Minimum slope upper bound
    DL_PD_SMP_LO   : TIME := T#10MS;         // 采样周期下限 / Sampling period lower bound
    DL_PD_SMP_HI   : TIME := T#1000MS;       // 采样周期上限 / Sampling period upper bound
    DL_PD_SEG_LO   : TIME := T#1S;           // 段超时下限 / Segment timeout lower bound
    DL_PD_SEG_HI   : TIME := T#1800S;        // 段超时上限 / Segment timeout upper bound
END_VAR

// 段 1｜输出与单拍标志预置
bProfileOk := FALSE;                                // 合格标志预清 / Acceptable flag pre-cleared
bSlowWarn := _bSlowLatch;                           // 早停建议由段内锁存派生（新循环起点即清） / Advice derived from the segment latch
eErr := 0;                                          // 错误码预清 / Error code pre-cleared

// 段 2｜采样与段超时定时器、沿实例无条件周期刷新
_tonSample(IN := bEnable AND bPumpOn AND (NOT _tonSample.Q), PT := tSampleTime);
_rtrigSample(CLK := _tonSample.Q);
_tonSeg(IN := bEnable AND bPumpOn AND (_eSeg <> E_DL_PumpSeg.eIdle) AND (_eSeg <> E_DL_PumpSeg.eDone)
            AND (_eSeg <> E_DL_PumpSeg.eFault), PT := tSegMax);

// 段 3｜首扫初始化（判据取非，R19）
IF NOT _bInit THEN
    _eSeg := E_DL_PumpSeg.eIdle;                    // 段待机起步 / Segment starts idle
    _bInit := TRUE;                                 // 首扫只做一次 / The first scan runs once
END_IF

// 段 4｜组态闸（段界反置使段永远进不去；最小抽速与采样周期判零防除零）
_bCfgOk := (fSeg1End_kPa > fSeg2End_kPa)
        AND NOT ((fSlopeMin_kPas <> fSlopeMin_kPas) OR ((fSlopeMin_kPas - fSlopeMin_kPas) <> (fSlopeMin_kPas - fSlopeMin_kPas)))
        AND (fSlopeMin_kPas >= DL_PD_SLOPE_LO) AND (fSlopeMin_kPas <= DL_PD_SLOPE_HI)
        AND (tSampleTime >= DL_PD_SMP_LO) AND (tSampleTime <= DL_PD_SMP_HI)
        AND (tSegMax >= DL_PD_SEG_LO) AND (tSegMax <= DL_PD_SEG_HI);
_fSampleSec := TIME_TO_LREAL(tSampleTime) / 1000.0; // 采样周期换算秒 [s] / Sampling period in seconds
IF _fSampleSec < 0.001 THEN
    _fSampleSec := 0.001;                           // 换算兜底下限 [s] / Conversion lower bound guard
END_IF
IF NOT _bCfgOk THEN
    eErr := DL_PD_CFG_BAD;                          // 故障级：组态非法 / Fault, bad configuration
    _uLatchCode := DL_PD_CFG_BAD;                   // 故障锁存码 / Fault latch code
    _eSeg := E_DL_PumpSeg.eFault;
END_IF

// 段 5｜压强可读闸（不可读不许推进段）
IF (fPress_kPa <> fPress_kPa) OR ((fPress_kPa - fPress_kPa) <> (fPress_kPa - fPress_kPa)) THEN
    eErr := DL_PD_PRESS_BAD;                        // 故障级：压强非有限 / Fault, the pressure is not finite
    _uLatchCode := DL_PD_PRESS_BAD;                 // 故障锁存码 / Fault latch code
    _eSeg := E_DL_PumpSeg.eFault;
    _bHasSample := FALSE;                           // 样本作废 / The sample is dropped
END_IF

// 段 6｜采样斜率（仅泵运行且样本有效）
IF _rtrigSample.Q AND _bHasSample AND (_eSeg <> E_DL_PumpSeg.eFault) THEN
    _fSlope := (fPress_kPa - _fPrev_kPa) / _fSampleSec;   // 本拍斜率（负 = 下降）[kPa/s] / Slope of this scan
    IF _eSeg = E_DL_PumpSeg.eRough THEN
        fSeg1Slope_kPas := ABS(_fSlope);            // 段 1 斜率取绝对值 [kPa/s] / Segment one slope magnitude
    ELSIF _eSeg = E_DL_PumpSeg.eTrans THEN
        fSeg2Slope_kPas := ABS(_fSlope);            // 段 2 斜率取绝对值 [kPa/s] / Segment two slope magnitude
    END_IF
    IF ABS(_fSlope) < fSlopeMin_kPas THEN
        _bSlowLatch := TRUE;                        // 低于包络：早停建议锁存 / Below the envelope, the advice is latched
        bSlowWarn := TRUE;
    END_IF
END_IF
IF _rtrigSample.Q THEN
    _fPrev_kPa := fPress_kPa;                       // 样本快照（唯一写点） / Sample snapshot, the single write point
    _bHasSample := TRUE;
END_IF

// 段 7｜段推进（ENUM + CASE + ELSE 兜底）
IF bEnable THEN
    CASE _eSeg OF
        E_DL_PumpSeg.eIdle:                         // 待机：泵启动即入粗抽
            IF bPumpOn THEN
                _bSlowLatch := FALSE;               // 新循环：建议清 / New cycle, the advice is cleared
                bSlowWarn := FALSE;                 // 同拍清出口，不留给上位幽灵建议 / The output is cleared in the same scan
                _bS1Judged := FALSE;
                _bS2Judged := FALSE;
                bProfileOk := FALSE;
                fSeg1Slope_kPas := 0.0;
                fSeg2Slope_kPas := 0.0;
                _eSeg := E_DL_PumpSeg.eRough;
            END_IF
            eErr := DL_PD_READY;

        E_DL_PumpSeg.eRough:                        // 粗抽段：跌破段界 1 即判段 1 合格与否
            IF NOT bPumpOn THEN
                _eSeg := E_DL_PumpSeg.eDone;        // 泵停：结束本次监视 / The pump stopped, the monitoring ends
            ELSIF fPress_kPa <= fSeg1End_kPa THEN
                IF ABS(fSeg1Slope_kPas) < fSlopeMin_kPas THEN
                    _bSlowLatch := TRUE;            // 段 1 低于包络 / Segment one below the envelope
                    bSlowWarn := TRUE;
                ELSE
                    _bS1Judged := TRUE;             // 段 1 合格 / Segment one accepted
                END_IF
                _eSeg := E_DL_PumpSeg.eTrans;
            ELSIF _tonSeg.Q THEN
                eErr := DL_PD_SEG_TO;               // 信息级：段超时，只建议早停 / Info, the segment timed out, advice only
                bSlowWarn := TRUE;
            END_IF

        E_DL_PumpSeg.eTrans:                        // 过渡段：跌破段界 2 即判段 2
            IF NOT bPumpOn THEN
                _eSeg := E_DL_PumpSeg.eDone;
            ELSIF fPress_kPa <= fSeg2End_kPa THEN
                IF ABS(fSeg2Slope_kPas) < fSlopeMin_kPas THEN
                    _bSlowLatch := TRUE;            // 段 2 低于包络 / Segment two below the envelope
                    bSlowWarn := TRUE;
                ELSE
                    _bS2Judged := TRUE;             // 段 2 合格 / Segment two accepted
                END_IF
                _eSeg := E_DL_PumpSeg.eFine;
            ELSIF _tonSeg.Q THEN
                eErr := DL_PD_SEG_TO;               // 信息级：段超时 / Info, the segment timed out
                bSlowWarn := TRUE;
            END_IF

        E_DL_PumpSeg.eFine:                         // 精抽段：泵停即完成并给全程结论
            IF NOT bPumpOn THEN
                bProfileOk := _bS1Judged AND _bS2Judged AND (NOT _bSlowLatch);   // 全程合格判据 / Whole-profile verdict
                _eSeg := E_DL_PumpSeg.eDone;
            ELSIF _tonSeg.Q THEN
                eErr := DL_PD_SEG_TO;               // 信息级：精抽段超时 / Info, the fine segment timed out
                bSlowWarn := TRUE;
            END_IF

        E_DL_PumpSeg.eDone:                         // 完成：等泵再次启动或失能
            bProfileOk := _bS1Judged AND _bS2Judged AND (NOT _bSlowLatch);
            IF NOT bPumpOn THEN
                _eSeg := E_DL_PumpSeg.eIdle;        // 泵已停：回待机 / Pump stopped, back to idle
            END_IF

        E_DL_PumpSeg.eFault:                        // 故障：停段，等失能后恢复
            IF _uLatchCode <> 0 THEN
                eErr := _uLatchCode;                // 锁存码回放（守住首因，不按当下输入改码） / Replay the latch code
            ELSIF eErr = 0 THEN
                eErr := DL_PD_PRESS_BAD;            // 兜底：无锁存码时按读数不可信上报 / Fallback when no latch code exists
            END_IF
            IF NOT bEnable THEN
                _eSeg := E_DL_PumpSeg.eIdle;        // 失能恢复 / Recovered on disable
                _uLatchCode := 0;                   // 锁存码清 / Latch code cleared
                _bHasSample := FALSE;
            END_IF

        ELSE
            // 非法段兜底（故障级，组态非法码承载）
            eErr := DL_PD_CFG_BAD;                  // 故障级：非法段值 / Fault, illegal segment value
            _uLatchCode := DL_PD_CFG_BAD;           // 故障锁存码 / Fault latch code
            _eSeg := E_DL_PumpSeg.eFault;
    END_CASE
END_IF

uSeg := 0;                                          // 段出口预置 / Segment output pre-set
CASE _eSeg OF
    E_DL_PumpSeg.eIdle:  uSeg := 0;                 // 待机 / Idle
    E_DL_PumpSeg.eRough: uSeg := 1;                 // 粗抽 / Rough
    E_DL_PumpSeg.eTrans: uSeg := 2;                 // 过渡 / Transition
    E_DL_PumpSeg.eFine:  uSeg := 3;                 // 精抽 / Fine
    E_DL_PumpSeg.eDone:  uSeg := 4;                 // 完成 / Done
    E_DL_PumpSeg.eFault: uSeg := 9;                 // 故障 / Fault
    ELSE
        uSeg := 9;                                  // 非法段按故障段出口 / Illegal segments are reported as fault
END_CASE
END_FUNCTION_BLOCK

(* ---- FB_DL_PvSoilingLossRate.st ---- *)
(*
  FB_DL_PvSoilingLossRate  —  组件积灰损失率估算与清洗提醒 / PV soiling loss estimation and cleaning reminder
  分类 Category : DL_Process
  码位 Code     : 16#06_0_85
  版本 Version  : 1.0.0
  溯源 Source   : LGF Measurement 语义借鉴 · clean-room 实现，仅借分类/参数域/命名，未复制源码
  功能 Function : 1) 仅在「辐照/温度同窗」条件下把性能比样本纳入基线窗口，避免把天气变化当积灰；
                  2) 用窗口均值作为基线、当前性能比相对基线的衰减速率按日折算；
                  3) 衰减速率分母（评估时间窗）先判正域；辐照低于下限时冻结估算并置 bFrozen，禁以低辐照数据外推。
  边界 Boundary : ① 基线在辐照/温度同窗条件下取，同窗外样本不纳入；
                  ② 衰减速率分母时间窗 > 0（防除零），非法即冻结；
                  ③ 辐照低于下限时冻结估算并置 bFrozen，禁低辐照外推；
                  ④ 结论态三行同向：性能比 → 基线 → 冻结/提醒标志。
  依赖 Depends  : FB_DL_SignalStatistics（基线窗口统计，每拍无条件调用）

  码表 Error codes（本件子码步进 16#10，避让邻件码位）:
    16#0002_0685 故障级：组态非法（辐照下限 <= 0 / 温度带宽 <= 0 / 评估时间窗 <= 0）
    16#0002_0695 故障级：窗口样本数为 0 却进入速率相（枚举/顺序兜底路径）
    16#0002_06A5 信息级：低辐照冻结估算（信息级，不置 bError）
*)

TYPE E_DL_PvSoilPhase :
(
    eIdle    := 0,   // 空闲 / Idle
    eCollect := 10,  // 同窗采样 / Same-window sampling
    eRate    := 20,  // 衰减速率计算 / Decay rate computation
    eAlarm   := 30,  // 清洗提醒 / Cleaning reminder
    eFrozen  := 40,  // 低辐照冻结 / Frozen at low irradiance
    eFault   := 90   // 故障锁定 / Fault locked
);
END_TYPE

FUNCTION_BLOCK FB_DL_PvSoilingLossRate
VAR_INPUT
    bEnable        : BOOL;                        // 总使能，FALSE 回空闲 / Master enable
    bSample        : BOOL := TRUE;                // 采样使能 / Sampling enable
    bReset         : BOOL;                        // 复位，上升沿清故障与统计窗 / Reset, clears fault and window
    fPowerKw       : REAL;                        // 组件实测输出功率 [kW]，域 > 0 / Measured module power [kW]
    fPowerRefKw    : REAL := 1.0;                 // 标称峰值功率 [kW]，域 > 0（性能比分母）/ Nameplate peak power [kW]
    fIrradWm2      : REAL;                        // 平面辐照度 [W/m2]，域 0~1500 / Plane-of-array irradiance [W/m2]
    fTempC         : REAL;                        // 组件背板温度 [degC]，域 −40~120 / Module back temperature [degC]
    fIrradMinWm2   : REAL := 400.0;               // 同窗辐照下限 [W/m2]，域 > 0 / Same-window irradiance floor
    fTempBandC     : REAL := 3.0;                 // 同窗温度带宽 [degC]，域 > 0 / Same-window temperature band
    fTempRefC      : REAL := 25.0;                // 同窗温度中心 [degC] / Same-window temperature centre
    fEvalSpanH     : REAL := 24.0;                // 评估时间窗 [h]，域 > 0（速率分母）/ Evaluation span [h]
    fLossAlarmPct  : REAL := 3.0;                 // 损失率清洗门限 [%]，域 0~100 / Soiling loss cleaning limit [%]
    nWindowLen     : INT := 32;                   // 基线窗口样本数 [个]，域 2~64 / Baseline window length
    fEps           : REAL := 1.0E-6;              // 浮点判零容差 [1] / Floating zero tolerance
END_VAR
VAR_OUTPUT
    fPrNowPct      : REAL;                        // 当前性能比 [%] / Current performance ratio [%]
    fPrBasePct     : REAL;                        // 基线性能比（窗口均值）[%] / Baseline performance ratio [%]
    fLossPct       : REAL;                        // 积灰损失率 [%] = (基线 − 当前) / 基线 × 100 / Soiling loss [%]
    fDecayPctPerDay : REAL;                       // 衰减速率 [%/天] / Decay rate [percent per day]
    bFrozen        : BOOL;                        // 估算冻结标志（保持型）/ Estimation frozen, held
    bCleanReminder : BOOL;                        // 清洗提醒（保持型）/ Cleaning reminder, held
    bError         : BOOL;                        // 故障标志，与故障级码配对 / Fault flag paired with fault codes
    uErrorId       : UDINT;                       // 事件码，0 = 无事件 / Event code, 0 = none
    eStateOut      : E_DL_PvSoilPhase;            // 状态机当前态，段尾单点映射 / Phase mapped at tail
END_VAR
VAR
    _eState        : E_DL_PvSoilPhase := E_DL_PvSoilPhase.eIdle;  // 内部状态 / Internal state
    rtrReset       : R_TRIG;                      // 复位沿 / Reset edge
    statPr         : FB_DL_SignalStatistics;      // 性能比窗口统计实例（无条件调用）/ PR window statistics
    bCfgOk         : BOOL;                        // 组态合法标志 / Configuration valid
    bWinOk         : BOOL;                        // 同窗条件满足标志 / Same-window condition met
    bIrradOk       : BOOL;                        // 辐照高于下限标志 / Irradiance above floor
    fPrPct         : REAL;                        // 性能比暂存 [%] / Performance ratio buffer [%]
    fLossBuf       : REAL;                        // 损失率暂存 [%] / Loss buffer [%]
    fSpanDay       : REAL;                        // 评估时间窗折算天数 [天] / Evaluation span in days
    uFault         : UDINT;                       // 锁存故障码 / Latched fault code
    uInfo          : UDINT;                       // 信息级码 / Information code
END_VAR
VAR CONSTANT
    DL_PV_PCTMAX   : REAL := 100.0;               // 百分比满量程 [%] / Full-scale percentage [%]
    DL_PV_HOURDAY  : REAL := 24.0;                // 每日小时数 [h] / Hours per day [h]
    DL_PV_IRRMAX   : REAL := 1500.0;              // 辐照物理域上限 [W/m2] / Irradiance domain high
END_VAR

(* === 段 0 · 实例刷新（无条件周期调用）=== *)
rtrReset(CLK := bReset);                          // 每拍刷新复位沿

(* === 段 1 · 组态闸与同窗判据 === *)
bCfgOk := (fPowerRefKw > fEps) AND (fIrradMinWm2 > fEps) AND (fTempBandC > fEps)
          AND (fEvalSpanH > fEps) AND (fPowerRefKw = fPowerRefKw)
          AND (fIrradMinWm2 = fIrradMinWm2) AND (fTempBandC = fTempBandC)
          AND (fEvalSpanH = fEvalSpanH);                          // 含 NaN 自反判据
IF NOT bCfgOk THEN
    uFault := 16#0002_0685;                       // 故障级：组态非法
END_IF
IF rtrReset.Q THEN
    uFault := 16#0000;                            // 复位沿清锁存（故障复位路径）
    bCleanReminder := FALSE;                      // 清洗提醒同步复位
END_IF
bIrradOk := (fIrradWm2 = fIrradWm2) AND (fIrradWm2 >= fIrradMinWm2)
            AND (fIrradWm2 <= DL_PV_IRRMAX);  // 辐照有限 + 高于同窗下限
bWinOk := bIrradOk
          AND (fTempC = fTempC) AND (ABS(fTempC - fTempRefC) <= fTempBandC)   // 温度同窗带宽
          AND (fPowerKw = fPowerKw) AND (fPowerKw > 0.0);                     // 功率正域闸（性能比分母）
IF bWinOk THEN
    fPrPct := fPowerKw / fPowerRefKw * DL_PV_PCTMAX;   // 性能比 [%]，分母已在组态闸判正
ELSE
    fPrPct := 0.0;                                // 同窗外不计性能比（0 仅作占位，样本不采样）
END_IF
fPrNowPct := fPrPct;                              // 当前性能比输出

(* === 段 2 · 基线窗口统计实例（每拍无条件调用）=== *)
statPr(fIn := fPrPct,                             // 输入当前性能比
       bSample := bWinOk AND bSample AND bCfgOk,  // 仅同窗样本纳入基线（防把天气当积灰）
       nWindow := nWindowLen,                     // 窗口长度，块内自钳 2~64
       bClear := rtrReset.Q);                     // 复位清窗
fPrBasePct := statPr.fMean;                       // 基线 = 窗口均值
fSpanDay := fEvalSpanH / DL_PV_HOURDAY;           // 时间窗折算天数，分母为正常量 24

(* === 段 3 · 主状态机（ENUM + CASE，含 ELSE 兜底）=== *)
CASE _eState OF
E_DL_PvSoilPhase.eIdle :
    bFrozen := FALSE;                             // 空闲不冻结
    uInfo := 16#0000;                             // 信息码清零
    IF uFault = 16#0002_0685 THEN
        _eState := E_DL_PvSoilPhase.eFault;       // 组态故障优先
    ELSIF bEnable AND bSample THEN
        _eState := E_DL_PvSoilPhase.eCollect;     // 进入采样相
    END_IF

E_DL_PvSoilPhase.eCollect :
    IF NOT bIrradOk THEN
        bFrozen := TRUE;                          // 低辐照：冻结估算，禁外推
        uInfo := 16#0002_06A5;                    // 信息级：低辐照冻结
        _eState := E_DL_PvSoilPhase.eFrozen;
    ELSIF (NOT statPr.bValid) OR (NOT statPr.bStatValid) THEN
        _eState := E_DL_PvSoilPhase.eCollect;     // 基线窗口未成形：继续采样（本拍不推进）
    ELSIF bCfgOk AND (fSpanDay > fEps) THEN
        _eState := E_DL_PvSoilPhase.eRate;        // 分母（时间窗）已判正，转速率相
    ELSE
        bFrozen := TRUE;                          // 分母非法：冻结
        _eState := E_DL_PvSoilPhase.eFrozen;
    END_IF

E_DL_PvSoilPhase.eRate :
    IF ABS(fPrBasePct) > fEps THEN                // 基线上分母防除零
        fLossBuf := (fPrBasePct - fPrPct) / fPrBasePct * DL_PV_PCTMAX;   // 积灰损失率
    ELSE
        fLossBuf := 0.0;                          // 基线近零：不出损失率（判不可测）
    END_IF
    IF fLossBuf < 0.0 THEN
        fLossBuf := 0.0;                          // 负损失（清洗后更干净）截零，不作负积灰显示
    END_IF
    IF fLossBuf > DL_PV_PCTMAX THEN
        fLossBuf := DL_PV_PCTMAX;                 // 饱和硬限（满量程 100%）
    END_IF
    fLossPct := fLossBuf;                         // 损失率输出
    fDecayPctPerDay := fLossBuf / fSpanDay;       // 衰减速率 [%/天]，分母已判 > fEps
    IF fLossBuf >= fLossAlarmPct THEN
        bCleanReminder := TRUE;                   // 置位型：清洗提醒（段尾不清零）
        _eState := E_DL_PvSoilPhase.eAlarm;
    ELSE
        bCleanReminder := FALSE;                  // 未达门限：提醒解除（可到达的解除路径）
        _eState := E_DL_PvSoilPhase.eCollect;
    END_IF

E_DL_PvSoilPhase.eAlarm :
    bCleanReminder := TRUE;                       // 提醒保持，等待清洗动作
    IF fLossPct < (fLossAlarmPct * 0.5) THEN
        bCleanReminder := FALSE;                  // 损失率降到门限一半以下：解除提醒
        _eState := E_DL_PvSoilPhase.eCollect;
    END_IF

E_DL_PvSoilPhase.eFrozen :
    bFrozen := TRUE;                              // 冻结标志保持
    IF bIrradOk AND bCfgOk AND statPr.bStatValid THEN
        bFrozen := FALSE;                         // 辐照恢复 + 窗口成形：解冻（可到达的解除路径）
        uInfo := 16#0000;                         // 信息码清除
        _eState := E_DL_PvSoilPhase.eCollect;
    END_IF

E_DL_PvSoilPhase.eFault :
    bFrozen := TRUE;                              // 故障态冻结估算
    fDecayPctPerDay := 0.0;                       // 速率输出 0（安全侧）
    IF uFault = 16#0000 THEN
        _eState := E_DL_PvSoilPhase.eIdle;        // 解锁后回空闲
    END_IF

ELSE
    _eState := E_DL_PvSoilPhase.eFault;           // 非法状态拦截
    uFault := 16#0002_0695;                       // 故障级：相 ID 越界（枚举兜底路径）
END_CASE
IF NOT bEnable THEN
    _eState := E_DL_PvSoilPhase.eIdle;            // 失能最高优先回空闲
    bFrozen := FALSE;                             // 失能不算冻结
    fDecayPctPerDay := 0.0;                       // 失能速率输出 0
END_IF

(* === 段 4 · 输出映射（三行同向：性能比 → 基线 → 标志）=== *)
IF NOT statPr.bStatValid THEN
    fDecayPctPerDay := 0.0;                       // 窗口未成形：速率不出结论
END_IF
bError := (uFault <> 16#0000);                    // 故障标志仅由故障级码置位（R45 配对）
IF bError THEN
    uErrorId := uFault;                           // 故障级优先上报
ELSE
    uErrorId := uInfo;                            // 否则上报信息级码
END_IF
eStateOut := _eState;                             // 输出枚举段尾单点映射（N2 规则）
END_FUNCTION_BLOCK
